(* IEC 61131-3 sources: plcassist-cli/packages/volt-lsp-iec/test-corpus/lenze-mid/Device/Plc Logic/Application/A70_MachineModuleSources/MM_MachineControl/01_Main, 9 files *)

(* ---- Mach1_Drives.fb ---- *)
FUNCTION_BLOCK Mach1_Drives
VAR_INPUT
END_VAR
VAR_OUTPUT
END_VAR
VAR
	testbyte: BYTE;
	testdint: DWORD;
	testword: WORD;
	OspRotationFlag: R_TRIG;
	OffDelayEnableDrivePower: TOF;
	EnableDrivePower: BOOL;
	bServoDrivesInSync: BOOL;
	TimeOutInSync: TON;
	bInSyncTimeOut: BOOL;
	TimeOutInLock: TON;
	tSetDrivesInLock: BOOL;
	bInLockTimeOut: BOOL;
	SideCorrection_CW: sUDT_ServoComm_Drive_Control;
	Servo_LimitJog_Instance: Servo_LimitJog;
	FBFeedforwardADS: FB_Lenze_i550;
	FBFeedforwardATF: FB_Lenze_i550;
	FBElevatorATF: FB_Lenze_i550;
	FBFan: FB_Lenze_i550;
	FBBobbin: FB_Lenze_i550;
	tReal: REAL;
	tWrapperStopPosition: DINT;

	sadad: FB_Lenze_i550;
	FB_Lenze_i550_0: FB_Lenze_i550;

mydword:DWORD;

	tbool: BOOL;
	OnDelayEnableSync: TON;
	ScaleBobbinTorque: LIN_TRAFO;
	tBobbinTorque: REAL;
	OffDelaySync: TOF;
	TON_0: TON;

	MainDrive_VirtualMasterControl: VirtualMasterControl;
END_VAR

VAR CONSTANT
	ctCurveIsSpeed: INT := 2;
	ctCurveIs0ToMax: INT := 0;
END_VAR
VAR
	ServoMainDrive: ServoControl;
	ServoWrappingDevice: ServoControl;
	ServoSideCorrection: ServoControl;
END_VAR

NETWORK 0 LD TITLE: "DONE network 3 : All drives ready"
  Mach1.GenFlags.ConditionsReadyForOperation := ((Mach1_Data.Drives.MainDrive.Status.DriveIsReady OR NOT Mach1_Data.Drives.MainDrive.Control.SetDriveEnable) AND (Mach1_Data.Drives.WrappingDevice.Status.DriveIsReady OR NOT Mach1_Data.Drives.WrappingDevice.Control.SetDriveEnable) AND (Mach1_Data.Drives.SideCorrection.Status.DriveIsReady OR NOT Mach1_Data.Drives.SideCorrection.Control.SetDriveEnable));
END_NETWORK
NETWORK 1 LD
  LET g24 := EnableDrivePower;
  Mach1_Data.Drives.WrappingDevice.Control.StartSetHomePos R= (g24 AND Mach1_Data.Drives.WrappingDevice.Status.DriveIsHomed);
  Mach1_Data.Drives.WrappingDevice.Control.StartSetHomePos S= ((g24 AND NOT Mach1_Data.Drives.WrappingDevice.Status.DriveIsHomed) AND FF500ms);
END_NETWORK
NETWORK 2 LD TITLE: "DONE Network 4: Enable drive power"
  // The off delay ensures that the drive can stop before the power is removed from the drive. The power must be removed from the drive before it goes to STO. If the power remains on during STO, the drive will generate an error.
  EnableDrivePower := (TRUE AND Mach1_Safety.Status.STO_OK);
END_NETWORK
NETWORK 3 LD
  Mach1_AuxData.AllDrivesHomed := Mach1_Data.Drives.MainDrive.Status.DriveIsHomed;
END_NETWORK
NETWORK 4 LD
  LET g0 := TRUE;
  Mach1_Data.Drives.MainDrive_VM.Control.SetDriveEnable := (g0 AND mach1.Genflags.DelayAfterSTO);
  Mach1_Data.Drives.MainDrive_VM.Control.ResetError := ((g0 AND NOT Mach1_Data.Drives.MainDrive_VM.Status.DriveIsReady) AND FF100ms);
  LET en1 := g0;
  IF en1 THEN MainDrive_VirtualMasterControl(iAcc := 600, iDec := 1800, ioVirtualMaster := Mach1_Data.Drives.MainDrive_VM, ioVirtualMasterCom := Data_Exchange_Motion.Servo_VirtualMaster); END_IF
  LET en2 := g0;
  IF en2 THEN HMI_Var.Mach1.ActualSpeed := MOVE(Mach1_Data.Drives.MainDrive_VM.Status.ActSpeed); END_IF
  LET en3 := en2;
  IF en3 THEN HMI_Var.Mach1.Position := MOVE(Mach1_Data.Drives.MainDrive_VM.Status.ActXPos); END_IF
END_NETWORK
NETWORK 5 LD TITLE: "Warning: machine in manual homing mode"
  Alarms_V5_1_100(Mach1_Alarms, (Mach1.GenFlags.DelayAfterSTO AND Mach1_AuxData.EnableManualHomeSetting), Mach1.GenFlags.ResetFlag, Mach1_Alarms.Alm033, Mach1.GenFlags.Warning);
END_NETWORK
NETWORK 6 LD TITLE: "DONE Network 5 : Conditions for sync/lock"
  LET g1 := Mach1.GenFlags.DelayAfterEmergStop;
  Mach1_AuxData.SetDrivesInSync := (TON_0(IN := (OffDelaySync(IN := (g1 AND Mach1_Safety.Status.DoorsOK), PT := T#500MS) AND Mach1_Safety.Status.STO_OK), PT := T#500MS) AND Mach1.GenFlags.ConditionsReadyForOperation AND Mach1_AuxData.AllDrivesHomed AND NOT Mach1_AuxData.EnableManualHomeSetting);
  LET g2 := (g1 AND Mach1_AuxData.SetDrivesInSync);
  bServoDrivesInSync := (g2 AND Mach1_Data.Drives.MainDrive.Status.InSync AND (Mach1_Data.Drives.WrappingDevice.Status.InSync OR NOT Mach1_Data.Drives.WrappingDevice.Control.SetDriveEnable) AND (Mach1_Data.Drives.SideCorrection.Status.InSync OR NOT Mach1_Data.Drives.SideCorrection.Control.SetDriveEnable));
  bInSyncTimeOut := TimeOutInSync(IN := (g2 AND NOT bServoDrivesInSync), PT := T#10S);
  Mach1_AuxData.SetDrivesInLock := ((g1 AND bServoDrivesInSync) AND (Mach1_AuxData.IEC_TIMERS.OffDelayLockDrives(IN := , PT := T#2s) OR TRUE));
  LET g3 := (g1 AND (Mach1_AuxData.SetDrivesInLock OR Mach1_AuxData.SetDrivesInSync));
  Mach1_AuxData.AllDrivesInLock := (g3 AND Mach1_Data.Drives.MainDrive.Status.InSync AND (Mach1_Data.Drives.WrappingDevice.Status.InSync OR NOT Mach1_Data.Drives.WrappingDevice.Control.SetDriveEnable) AND (Mach1_Data.Drives.SideCorrection.Status.InSync OR NOT Mach1_Data.Drives.SideCorrection.Control.SetDriveEnable));
  bInLockTimeOut := TimeOutInLock(IN := (g3 AND NOT Mach1_AuxData.AllDrivesInLock), PT := T#5S);
  tSetDrivesInLock := g3;
END_NETWORK
NETWORK 7 LD TITLE: "DONE Network 6: Servo Main drive: Control"
  LET g4 := TRUE;
  Mach1_Data.Drives.MainDrive_VM.Control.StartMovement := (g4 AND ((Mach1_Safety.Control.RequestManSpeed AND Mach1_Safety.Status.SafetyManSpeed) OR (Mach1_Safety.Control.RequestAutoSpeed AND Mach1_Safety.Status.SafetyAutoSpeed)));
  LET en1 := (g4 AND TRUE);
  IF en1 THEN Mach1_Data.Drives.MainDrive.CAM.CamType := MOVE(ctCurveIs0ToMax); END_IF
  Mach1_Data.Drives.MainDrive.Control.SetInSync := (en1 AND tSetDrivesInLock);
  LET g5 := (g4 AND TRUE);
  Mach1_Data.Drives.MainDrive.Control.SetBrakeRelease := (g5 AND Mach1_Alarms.Alm001 AND HMI_Var.ReleaseBrake);
  HMI_Var.ReleaseBrake R= (g5 AND (NOT Mach1_Alarms.Alm001 OR (mach1.Genflags.StartFlag AND Mach1_Alarms.Alm001)));
  LET en2 := (g4 AND TRUE);
  IF en2 THEN ServoMainDrive(iServoStatus := Data_Exchange_Motion.Servo_MainDrive.Status, iEnableHomeMovement := TRUE, iEnablePower := EnableDrivePower, iFF100ms := LST_General.FF100ms, ioUDT_ServoDrive := Mach1_Data.Drives.MainDrive, oServoControl => Data_Exchange_Motion.Servo_MainDrive.Control); END_IF
  Mach1.GenFlags.Rotflag := OspRotationFlag(CLK := (en2 AND Mach1_Data.Drives.MainDrive.Status.RotationPulse));
END_NETWORK
NETWORK 8 LD TITLE: "DONE Network 7 : Servo Main drive: Alarms"
  Mach1.GenFlags.StopDriveDirect S= (Alarms_V5_1_100(Mach1_Alarms, (Mach1.GenFlags.DelayAfterSTO AND NOT Mach1_Data.Drives.MainDrive.Status.DriveIsReady), Mach1.GenFlags.ResetFlag, Mach1_Alarms.Alm020, Mach1.GenFlags.MinorAlarm) OR Alarms_V5_1_100(Mach1_Alarms, (Mach1.GenFlags.DelayAfterSTO AND Mach1_Data.Drives.MainDrive.Status.DriveTorqueError), Mach1.GenFlags.ResetFlag, Mach1_Alarms.Alm021, Mach1.GenFlags.MinorAlarm) OR Alarms_V5_1_100(Mach1_Alarms, (Mach1.GenFlags.DelayAfterSTO AND NOT Mach1_Data.Drives.MainDrive.Status.DriveIsHomed), Mach1.GenFlags.ResetFlag, Mach1_Alarms.Alm022, Mach1.GenFlags.MinorAlarm));
END_NETWORK
NETWORK 9 LD
  Mach1_Data.Drives.MainDrive.Control.ResetError S= (((Mach1_Alarms.Alm020 OR Mach1_Alarms.Alm021 OR Mach1_Alarms.Alm022) AND Mach1.GenFlags.ResetFlag) OR (TON_0.Q AND Imp100ms AND Mach1_Safety.Status.ServiceMode AND Mach1_Safety.Status.Service_ButtonAB));
END_NETWORK
NETWORK 10 LD TITLE: "DONE Network 8: Servo Wrapping device: Control"
  LET g6 := TRUE;
  LET en1 := (g6 AND TRUE);
  IF en1 THEN Mach1_Data.Drives.WrappingDevice.CAM.CamType := MOVE(ctCurveIsSpeed); END_IF
  Mach1_Data.Drives.WrappingDevice.Control.SetInSync := (en1 AND tSetDrivesInLock);
  LET en2 := g6;
  IF en2 THEN Mach1_Data.Drives.WrappingDevice.CAM.Y_Scale_Recipe := MOVE(Mach1_Data.Settings.Ints.RollingDeviceSpeedFactor); END_IF
  LET en3 := (g6 AND TRUE);
  IF en3 THEN ServoWrappingDevice(iServoStatus := Data_Exchange_Motion.Servo_WrappingDevice.Status, iEnableHomeMovement := TRUE, iEnablePower := EnableDrivePower, iFF100ms := LST_General.FF100ms, ioUDT_ServoDrive := Mach1_Data.Drives.WrappingDevice, oServoControl => Data_Exchange_Motion.Servo_WrappingDevice.Control); END_IF
END_NETWORK
NETWORK 11 LD TITLE: "DONE Network 9 : Servo Wrapping Device: Alarms"
  LET g7 := (Alarms_V5_1_100(Mach1_Alarms, (Mach1.GenFlags.DelayAfterSTO AND NOT Mach1_Data.Drives.WrappingDevice.Status.DriveIsReady AND Mach1_Data.Drives.WrappingDevice.Control.SetDriveEnable), Mach1.GenFlags.ResetFlag, Mach1_Alarms.Alm023, Mach1.GenFlags.MinorAlarm) OR Alarms_V5_1_100(Mach1_Alarms, (Mach1.GenFlags.DelayAfterSTO AND Mach1_Data.Drives.WrappingDevice.Status.DriveTorqueError), Mach1.GenFlags.ResetFlag, Mach1_Alarms.Alm024, Mach1.GenFlags.MinorAlarm) OR Alarms_V5_1_100(Mach1_Alarms, (Mach1.GenFlags.DelayAfterSTO AND NOT Mach1_Data.Drives.WrappingDevice.Status.DriveIsHomed), Mach1.GenFlags.ResetFlag, Mach1_Alarms.Alm025, Mach1.GenFlags.MinorAlarm));
  Mach1.GenFlags.StopDriveDirect S= g7;
  Mach1_Data.Drives.WrappingDevice.Control.ResetError S= (g7 AND Mach1.GenFlags.ResetFlag);
END_NETWORK
NETWORK 12 LD
  Mach1_Data.Drives.WrappingDevice.Control.ResetError S= (((Mach1_Alarms.Alm023 OR Mach1_Alarms.Alm024 OR Mach1_Alarms.Alm025) AND Mach1.GenFlags.ResetFlag) OR (TON_0.Q AND Imp100ms AND Mach1_Safety.Status.ServiceMode AND Mach1_Safety.Status.Service_ButtonAB));
END_NETWORK
NETWORK 13 LD
END_NETWORK
NETWORK 14 LD TITLE: "Digital inputs"
  // 16: non-motor side
  // 17: motor side
  LET en1 := TRUE;
  IF en1 THEN mydword := MOVE(%ID79); END_IF
  LET g8 := en1;
  Data_Exchange_Motion.Servo_SideCorrection.Status.Spare1 := (g8 AND mydword.16);
  Data_Exchange_Motion.Servo_SideCorrection.Status.Spare2 := (g8 AND mydword.17);
END_NETWORK
NETWORK 15 LD TITLE: "DONE Network 10: Servo Side correction: Control"
  LET g9 := TRUE;
  LET en1 := (g9 AND TRUE);
  IF en1 THEN Mach1_Data.Drives.SideCorrection.CAM.CamType := MOVE(ctCurveIsSpeed); END_IF
  Mach1_Data.Drives.SideCorrection.Control.SetInSync := (en1 AND tSetDrivesInLock);
  LET en2 := (g9 AND TRUE);
  IF en2 THEN ServoSideCorrection(iServoStatus := Data_Exchange_Motion.Servo_SideCorrection.Status, iEnableHomeMovement := TRUE, iEnablePower := EnableDrivePower, iFF100ms := LST_General.FF100ms, ioUDT_ServoDrive := Mach1_Data.Drives.SideCorrection, oServoControl => SideCorrection_CW); END_IF
  LET en3 := (g9 AND TRUE);
  IF en3 THEN Servo_LimitJog_Instance(iServoStatus := Data_Exchange_Motion.Servo_SideCorrection.Status, iServoControl := SideCorrection_CW, ioUDT_ServoDrive := Mach1_Data.Drives.SideCorrection, ioUDT_JogLimitFree := Mach1_Data.Drives.SideCorrection_FreeLimit, oServoControl => Data_Exchange_Motion.Servo_SideCorrection.Control); END_IF
END_NETWORK
NETWORK 16 LD TITLE: "DONE Network 11 : Servo Side correction: Alarms"
  LET g10 := (Alarms_V5_1_100(Mach1_Alarms, (Mach1.GenFlags.DelayAfterSTO AND NOT Mach1_Data.Drives.SideCorrection.Status.DriveIsReady AND Mach1_Data.Drives.SideCorrection.Control.SetDriveEnable), Mach1.GenFlags.ResetFlag, Mach1_Alarms.Alm026, Mach1.GenFlags.MinorAlarm) OR Alarms_V5_1_100(Mach1_Alarms, (Mach1.GenFlags.DelayAfterSTO AND Mach1_Data.Drives.SideCorrection.Status.DriveTorqueError), Mach1.GenFlags.ResetFlag, Mach1_Alarms.Alm027, Mach1.GenFlags.MinorAlarm) OR Alarms_V5_1_100(Mach1_Alarms, (Mach1.GenFlags.DelayAfterSTO AND NOT Mach1_Data.Drives.SideCorrection.Status.DriveIsHomed), Mach1.GenFlags.ResetFlag, Mach1_Alarms.Alm028, Mach1.GenFlags.MinorAlarm));
  Mach1.GenFlags.StopDriveDirect S= g10;
  Mach1_Data.Drives.SideCorrection.Control.ResetError S= (g10 AND Mach1.GenFlags.ResetFlag);
END_NETWORK
NETWORK 17 LD
  Mach1_Data.Drives.SideCorrection.Control.ResetError S= (((Mach1_Alarms.Alm026 OR Mach1_Alarms.Alm027 OR Mach1_Alarms.Alm028) AND Mach1.GenFlags.ResetFlag) OR (TON_0.Q AND Imp100ms AND Mach1_Safety.Status.ServiceMode AND Mach1_Safety.Status.Service_ButtonAB));
END_NETWORK
NETWORK 18 LD
END_NETWORK
NETWORK 19 LD TITLE: "DONE Network 12: Feedforward ADS"
  LET g11 := TRUE;
  Mach1_Data.Drives.FeedForwardADS.Control.Enable := (g11 AND Mach1.GenFlags.DelayAfterEmergStop AND NOT Mach1_Alarms.Alm015);
  Mach1_Data.Drives.FeedForwardADS.Control.Reverse := g11;
  LET en1 := g11;
  IF en1 THEN FBFeedforwardADS(iStatusWord := Data_Exchange_Motion.FQI_FeedforwardADS.Status, iGearRatioNumerator := 2790.0, iGearRatioDenominator := 111.0, iNominalMotorSpeedwoSlipComp_RPM := 3000.0, iNominalMotorFrequency_Hz := 100.0, iAxisJogSpeed_RPM := 10.0, ioUDT := Mach1_Data.Drives.FeedForwardADS, oControlWord => Data_Exchange_Motion.FQI_FeedforwardADS.Controlword, oRefSpeed => Data_Exchange_Motion.FQI_FeedforwardADS.RefSpeed); END_IF
END_NETWORK
NETWORK 20 LD TITLE: "DONE Network 13: Alarms feed forward dryer"
  LET g12 := Alarms_V5_1_100(Mach1_Alarms, (Mach1.GenFlags.DelayAfterEmergStop AND Mach1_Data.Drives.FeedForwardADS.Status.Error), True, Mach1_Alarms.Alm015, Mach1.GenFlags.MinorAlarm);
  Mach1.GenFlags.StopDriveDirect S= g12;
  Mach1_Data.Drives.FeedForwardADS.Control.ResetError S= (g12 AND Mach1.GenFlags.ResetFlag);
END_NETWORK
NETWORK 21 LD TITLE: "DONE Network 14: Feedforward ATF"
  LET g13 := TRUE;
  Mach1_Data.Drives.FeedForwardATF.Control.Enable := (g13 AND Mach1.GenFlags.DelayAfterEmergStop AND NOT Mach1_Alarms.Alm016);
  LET en1 := g13;
  IF en1 THEN FBFeedforwardATF(iStatusWord := Data_Exchange_Motion.FQI_FeedforwardATF.Status, iGearRatioNumerator := 2790.0, iGearRatioDenominator := 111.0, iNominalMotorSpeedwoSlipComp_RPM := 3000.0, iNominalMotorFrequency_Hz := 100.0, iAxisJogSpeed_RPM := 10.0, ioUDT := Mach1_Data.Drives.FeedForwardATF, oControlWord => Data_Exchange_Motion.FQI_FeedforwardATF.Controlword, oRefSpeed => Data_Exchange_Motion.FQI_FeedforwardATF.RefSpeed); END_IF
END_NETWORK
NETWORK 22 LD TITLE: "DONE Network 15: Alarms feed forward trayfiller"
  LET g14 := Alarms_V5_1_100(Mach1_Alarms, (Mach1.GenFlags.DelayAfterEmergStop AND Mach1_Data.Drives.FeedForwardATF.Status.Error), True, Mach1_Alarms.Alm016, Mach1.GenFlags.MinorAlarm);
  Mach1.GenFlags.StopDriveDirect S= g14;
  Mach1_Data.Drives.FeedForwardATF.Control.ResetError S= (g14 AND Mach1.GenFlags.ResetFlag);
END_NETWORK
NETWORK 23 LD TITLE: "DONE Network 16: Elevator ATF"
  LET g15 := TRUE;
  Mach1_Data.Drives.ElevatorATF.Control.Enable := (g15 AND Mach1.GenFlags.DelayAfterEmergStop AND NOT Mach1_Alarms.Alm014);
  LET en1 := g15;
  IF en1 THEN FBElevatorATF(iStatusWord := Data_Exchange_Motion.FQI_ElevatorATF.Status, iGearRatioNumerator := 100.0, iGearRatioDenominator := 111.0, iNominalMotorSpeedwoSlipComp_RPM := 3000.0, iNominalMotorFrequency_Hz := 100.0, iAxisJogSpeed_RPM := 10.0, ioUDT := Mach1_Data.Drives.ElevatorATF, oControlWord => Data_Exchange_Motion.FQI_ElevatorATF.Controlword, oRefSpeed => Data_Exchange_Motion.FQI_ElevatorATF.RefSpeed); END_IF
END_NETWORK
NETWORK 24 LD TITLE: "DONE Network 17: Alarms Elevator trayfiller"
  LET g16 := Alarms_V5_1_100(Mach1_Alarms, (Mach1.GenFlags.DelayAfterEmergStop AND Mach1_Data.Drives.ElevatorATF.Status.Error), True, Mach1_Alarms.Alm014, Mach1.GenFlags.MinorAlarm);
  Mach1.GenFlags.StopDriveDirect S= g16;
  Mach1_Data.Drives.ElevatorATF.Control.ResetError S= (g16 AND Mach1.GenFlags.ResetFlag);
END_NETWORK
NETWORK 25 LD TITLE: "DONE Network 18: Fan"
  LET g26 := TRUE;
  Mach1_Data.Drives.Fan.Control.Enable := (g26 AND Mach1.GenFlags.EnableAuxDrive AND NOT Mach1_Alarms.Alm017);
  LET en1 := g26;
  IF en1 THEN FBFan(iStatusWord := Data_Exchange_Motion.FQI_Fan.Status, iGearRatioNumerator := 1.0, iGearRatioDenominator := 1.0, iNominalMotorSpeedwoSlipComp_RPM := 3000.0, iNominalMotorFrequency_Hz := 50.0, iAxisJogSpeed_RPM := 10.0, ioUDT := Mach1_Data.Drives.Fan, oControlWord => Data_Exchange_Motion.FQI_Fan.Controlword, oRefSpeed => Data_Exchange_Motion.FQI_Fan.RefSpeed); END_IF
END_NETWORK
NETWORK 26 LD TITLE: "DONE Network 19: Alarms Fan"
  LET g18 := Alarms_V5_1_100(Mach1_Alarms, (Mach1.GenFlags.DelayAfterEmergStop AND Mach1_Data.Drives.Fan.Status.Error), True, Mach1_Alarms.Alm017, Mach1.GenFlags.MinorAlarm);
  Mach1.GenFlags.StopDriveDirect S= g18;
  Mach1_Data.Drives.Fan.Control.ResetError S= (g18 AND Mach1.GenFlags.ResetFlag);
END_NETWORK
NETWORK 27 LD TITLE: "DONE Network 20: Bobbin"
  LET g19 := TRUE;
  LET en1 := (g19 AND Mach1.GenFlags.EnableAuxDrive AND NOT HMI_Var.Btn_Cleaning);
  IF en1 THEN (Mach1_Data.Settings.Ints.TorqueControlBobbin > 0); END_IF
  LET g20 := (en1 AND Mach1_Safety.Status.AllDoorsActuallyClosed);
  Mach1_Data.Drives.Bobbine.Control.Enable := g20;
  LET en2 := g20;
  IF en2 THEN Mach1_Data.Drives.Bobbine.Control.AutoSpeed := MOVE(860); END_IF
  Mach1_Data.Drives.Bobbine.Control.StartAuto := en2;
  LET en3 := g19;
  IF en3 THEN FBBobbin(iStatusWord := Data_Exchange_Motion.FQI_Bobbin.Status, iGearRatioNumerator := 2790.0, iGearRatioDenominator := 111.0, iNominalMotorSpeedwoSlipComp_RPM := 3000.0, iNominalMotorFrequency_Hz := 50.0, iAxisJogSpeed_RPM := 10.0, ioUDT := Mach1_Data.Drives.Bobbine, oControlWord => Data_Exchange_Motion.FQI_Bobbin.Controlword, oRefSpeed => Data_Exchange_Motion.FQI_Bobbin.RefSpeed); END_IF
  LET g21 := (g19 AND HMI_Var.Mach1.CalibrateTorqueValues);
  LET en4 := g21;
  IF en4 THEN Data_Exchange_Motion.BobbinTorque := MOVE(Mach1_AuxData.TorqueCalibrationValue); END_IF
  LET en5 := (g21 AND HMI_Var.Mach1.setMinTorqueValue);
  IF en5 THEN Mach1_Data.Settings.Dints.minTorqueValue := MOVE(Mach1_AuxData.TorqueCalibrationValue); END_IF
  HMI_Var.Mach1.setMinTorqueValue R= en5;
  LET en6 := (g21 AND HMI_Var.Mach1.setMaxTorqueValue);
  IF en6 THEN Mach1_Data.Settings.Dints.maxTorqueValue := MOVE(Mach1_AuxData.TorqueCalibrationValue); END_IF
  HMI_Var.Mach1.setMaxTorqueValue R= en6;
  LET i1 := DINT_TO_REAL(Mach1_Data.Settings.Dints.minTorqueValue);
  LET i2 := DINT_TO_REAL(Mach1_Data.Settings.Dints.maxTorqueValue);
  LET en7 := (g19 AND NOT HMI_Var.Mach1.CalibrateTorqueValues);
  IF en7 THEN ScaleBobbinTorque(IN := Mach1_Data.Settings.Ints.TorqueControlBobbin, IN_MIN := 0, IN_MAX := 1000, OUT_MIN := i1, OUT_MAX := i2, OUT => tBobbinTorque); END_IF
  LET i3 := REAL_TO_DINT(tBobbinTorque);
  LET en8 := en7;
  IF en8 THEN Data_Exchange_Motion.BobbinTorque := MOVE(i3); END_IF
END_NETWORK
NETWORK 28 LD TITLE: "DONE Network 21: Alarms Bobbine"
  LET g22 := Alarms_V5_1_100(Mach1_Alarms, (Mach1_AuxData.MIDS_Active AND Mach1.GenFlags.DelayAfterEmergStop AND NOT Mach1_Data.Drives.Bobbine.Status.DriveReady AND Mach1_AuxData.AllDrivesHomed), True, Mach1_Alarms.Alm010, Mach1.GenFlags.MinorAlarm);
  Mach1.GenFlags.StopDriveDirect S= g22;
  Mach1_Data.Drives.Bobbine.Control.ResetError S= (g22 AND Mach1.GenFlags.ResetFlag);
END_NETWORK
NETWORK 29 LD TITLE: "TODO Network 22:"
  // WRAPPER
END_NETWORK
NETWORK 30 LD TITLE: "TODO Network 23: Limit Wrapper stop position"
  LET g23 := TRUE;
  LET en1 := g23;
  IF en1 THEN (Mach1_Data.Settings.Dints.WrapperStopPosition > 400); END_IF
  LET en2 := en1;
  IF en2 THEN Mach1_Data.Settings.Dints.WrapperStopPosition := MOVE(400); END_IF
  LET en3 := g23;
  IF en3 THEN (Mach1_Data.Settings.Dints.WrapperStopPosition < 5); END_IF
  LET en4 := en3;
  IF en4 THEN Mach1_Data.Settings.Dints.WrapperStopPosition := MOVE(5); END_IF
  LET en5 := g23;
  IF en5 THEN tWrapperStopPosition := (Mach1_Data.Settings.Dints.WrapperStopPosition * 100); END_IF
END_NETWORK
NETWORK 31 LD TITLE: "TODO Network 25:"
  Data_Exchange_Motion.FeedForwardWrapper.Control.Enable := (TRUE AND Mach1.GenFlags.DelayAfterEmergStop AND NOT Mach1_Alarms.Alm066);
END_NETWORK
NETWORK 32 LD TITLE: "TODO Network 26:"
  LET g1 := (Alarms_V5_1_100(Mach1_Alarms, (Mach1_AuxData.MIDS_Active AND Mach1.GenFlags.EnableMainDrive AND HMI_Var.Test_Prod AND NOT HMI_Var.Btn_Cleaning AND Mach1_AuxData.AllDrivesHomed AND NOT Data_Exchange_Motion.FeedForwardWrapper.Status.ReadyForMotion), Mach1.Genflags.StartFlag, Mach1_Alarms.Alm056, Mach1.GenFlags.MinorAlarm) AND mach1.Genflags.ResetFlag);
  Mach1_Data.Drives.WrappingDevice.Control.ResetError S= g1;
  Data_Exchange_Motion.FeedForwardWrapper.Control.ResetError := g1;
END_NETWORK
NETWORK 33 LD TITLE: "TODO Network 27:"
  ;
END_NETWORK

END_FUNCTION_BLOCK

(* ---- fc_Information.prg ---- *)
PROGRAM fc_Information
VAR
END_VAR

VersionInfo_DB.PLC_version:='MID-S100-L-V00_00';
VersionInfo_DB.PLC_Version_Date:='08-06-2023';

END_PROGRAM

(* ---- ForceOutput.prg ---- *)
PROGRAM ForceOutput
VAR
END_VAR

NETWORK 0 LD
  LET g2 := HMI_Var.ForceOutputs;
  LST_InputsOutputs.Q100_0_Pilot_light_Alarm_green_ := (g2 AND LST_InputsOutputs.Serv_QB100.0);
  LST_InputsOutputs.Q100_1_Pilot_light_Alarm_orange_ := (g2 AND LST_InputsOutputs.Serv_QB100.1);
  LST_InputsOutputs.Q100_2_Pilot_light_Alarm_red_ := (g2 AND LST_InputsOutputs.Serv_QB100.2);
  LST_InputsOutputs.Q100_3_Pilot_light_Alarm_buzzer_ := (g2 AND LST_InputsOutputs.Serv_QB100.3);
  LST_InputsOutputs.Q100_4_Spare := (g2 AND LST_InputsOutputs.Serv_QB100.4);
  LST_InputsOutputs.Q100_5_Signal_lamp_Start := (g2 AND LST_InputsOutputs.Serv_QB100.5);
  LST_InputsOutputs.Q100_6_Signal_lamp_Stop := (g2 AND LST_InputsOutputs.Serv_QB100.6);
  LST_InputsOutputs.Q100_7_Activate_greasing_system := (g2 AND LST_InputsOutputs.Serv_QB100.7);
  LST_InputsOutputs.Q101_0_REL_release_brake := (g2 AND LST_InputsOutputs.Serv_QB101.0);
  LST_InputsOutputs.Q101_1_PNV_Waterlevel_control := (g2 AND LST_InputsOutputs.Serv_QB101.1);
  LST_InputsOutputs.Q101_2_Enable_GluePump := (g2 AND LST_InputsOutputs.Serv_QB101.2);
  LST_InputsOutputs.Q101_3_Spare := (g2 AND LST_InputsOutputs.Serv_QB101.3);
  LST_InputsOutputs.Q101_4_Spare := (g2 AND LST_InputsOutputs.Serv_QB101.4);
  LST_InputsOutputs.Q101_5_Spare := (g2 AND LST_InputsOutputs.Serv_QB101.5);
  LST_InputsOutputs.Q101_6_Spare := (g2 AND LST_InputsOutputs.Serv_QB101.6);
  LST_InputsOutputs.Q101_7_Spare := (g2 AND LST_InputsOutputs.Serv_QB101.7);
END_NETWORK
NETWORK 1 LD
  LET g1 := HMI_Var.ForceOutputs;
  LST_InputsOutputs.Q132_0_SL_Start_OP2a := (g1 AND LST_InputsOutputs.Serv_QB132.0);
  LST_InputsOutputs.Q132_1_SL_Stop_OP2a := (g1 AND LST_InputsOutputs.Serv_QB132.1);
  LST_InputsOutputs.Q132_2_Enable_power_controllers := (g1 AND LST_InputsOutputs.Serv_QB132.2);
  LST_InputsOutputs.Q132_3_Spare := (g1 AND LST_InputsOutputs.Serv_QB132.3);
  LST_InputsOutputs.Q132_4_CT_Fan_dryer := (g1 AND LST_InputsOutputs.Serv_QB132.4);
  LST_InputsOutputs.Q132_5_Spare := (g1 AND LST_InputsOutputs.Serv_QB132.5);
  LST_InputsOutputs.Q132_6_PNV_Inpusher := (g1 AND LST_InputsOutputs.Serv_QB132.6);
  LST_InputsOutputs.Q132_7_PNV_tilting_inpusher := (g1 AND LST_InputsOutputs.Serv_QB132.7);
  LST_InputsOutputs.Q133_0_Spare := (g1 AND LST_InputsOutputs.Serv_QB133.0);
  LST_InputsOutputs.Q133_1_Spare := (g1 AND LST_InputsOutputs.Serv_QB133.1);
  LST_InputsOutputs.Q133_2_Spare := (g1 AND LST_InputsOutputs.Serv_QB133.2);
  LST_InputsOutputs.Q133_3_Spare := (g1 AND LST_InputsOutputs.Serv_QB133.3);
  LST_InputsOutputs.Q133_4_Spare := (g1 AND LST_InputsOutputs.Serv_QB133.4);
  LST_InputsOutputs.Q133_5_InfeedConv_Fwd := (g1 AND LST_InputsOutputs.Serv_QB133.5);
  LST_InputsOutputs.Q133_6_InfeedConv_Rev := (g1 AND LST_InputsOutputs.Serv_QB133.6);
  LST_InputsOutputs.Q133_7_OutfeedConv_Fwd := (g1 AND LST_InputsOutputs.Serv_QB133.7);
END_NETWORK
NETWORK 2 LD
  LET g0 := HMI_Var.ForceOutputs;
  LST_InputsOutputs.Q136_0_Spare := (g0 AND LST_InputsOutputs.Serv_QB136.0);
  LST_InputsOutputs.Q136_1_Spare := (g0 AND LST_InputsOutputs.Serv_QB136.1);
  LST_InputsOutputs.Q136_2_Spare := (g0 AND LST_InputsOutputs.Serv_QB136.2);
  LST_InputsOutputs.Q136_3_Spare := (g0 AND LST_InputsOutputs.Serv_QB136.3);
  LST_InputsOutputs.Q136_4_Spare := (g0 AND LST_InputsOutputs.Serv_QB136.4);
  LST_InputsOutputs.Q136_5_Spare := (g0 AND LST_InputsOutputs.Serv_QB136.5);
  LST_InputsOutputs.Q136_6_Spare := (g0 AND LST_InputsOutputs.Serv_QB136.6);
  LST_InputsOutputs.Q136_7_Spare := (g0 AND LST_InputsOutputs.Serv_QB132.7);
  LST_InputsOutputs.Q137_0_Spare := (g0 AND LST_InputsOutputs.Serv_QB137.0);
  LST_InputsOutputs.Q137_1_Spare := (g0 AND LST_InputsOutputs.Serv_QB137.1);
  LST_InputsOutputs.Q137_2_Spare := (g0 AND LST_InputsOutputs.Serv_QB137.2);
  LST_InputsOutputs.Q137_3_Spare := (g0 AND LST_InputsOutputs.Serv_QB137.3);
  LST_InputsOutputs.Q137_4_Spare := (g0 AND LST_InputsOutputs.Serv_QB137.4);
  LST_InputsOutputs.Q137_5_Spare := (g0 AND LST_InputsOutputs.Serv_QB137.5);
  LST_InputsOutputs.Q137_6_Spare := (g0 AND LST_InputsOutputs.Serv_QB137.6);
  LST_InputsOutputs.Q137_7_Spare := (g0 AND LST_InputsOutputs.Serv_QB137.7);
END_NETWORK
NETWORK 3 LD
END_NETWORK

END_PROGRAM

(* ---- ForceOutput_1.prg ---- *)
PROGRAM ForceOutput_1
VAR
END_VAR

NETWORK 0 LD
  LET g2 := NOT HMI_Var.ForceOutputs;
  LST_InputsOutputs.Serv_QB100.0 := (g2 AND LST_InputsOutputs.Q100_0_Pilot_light_Alarm_green_);
  LST_InputsOutputs.Serv_QB100.1 := (g2 AND LST_InputsOutputs.Q100_1_Pilot_light_Alarm_orange_);
  LST_InputsOutputs.Serv_QB100.2 := (g2 AND LST_InputsOutputs.Q100_2_Pilot_light_Alarm_red_);
  LST_InputsOutputs.Serv_QB100.3 := (g2 AND LST_InputsOutputs.Q100_3_Pilot_light_Alarm_buzzer_);
  LST_InputsOutputs.Serv_QB100.4 := (g2 AND LST_InputsOutputs.Q100_4_Spare);
  LST_InputsOutputs.Serv_QB100.5 := (g2 AND LST_InputsOutputs.Q100_5_Signal_lamp_Start);
  LST_InputsOutputs.Serv_QB100.6 := (g2 AND LST_InputsOutputs.Q100_6_Signal_lamp_Stop);
  LST_InputsOutputs.Serv_QB100.7 := (g2 AND LST_InputsOutputs.Q100_7_Activate_greasing_system);
  LST_InputsOutputs.Serv_QB101.0 := (g2 AND LST_InputsOutputs.Q101_0_REL_release_brake);
  LST_InputsOutputs.Serv_QB101.1 := (g2 AND LST_InputsOutputs.Q101_1_PNV_Waterlevel_control);
  LST_InputsOutputs.Serv_QB101.2 := (g2 AND LST_InputsOutputs.Q101_2_Enable_GluePump);
  LST_InputsOutputs.Serv_QB101.3 := (g2 AND LST_InputsOutputs.Q101_3_Spare);
  LST_InputsOutputs.Serv_QB101.4 := (g2 AND LST_InputsOutputs.Q101_4_Spare);
  LST_InputsOutputs.Serv_QB101.5 := (g2 AND LST_InputsOutputs.Q101_5_Spare);
  LST_InputsOutputs.Serv_QB101.6 := (g2 AND LST_InputsOutputs.Q101_6_Spare);
  LST_InputsOutputs.Serv_QB101.7 := (g2 AND LST_InputsOutputs.Q101_7_Spare);
END_NETWORK
NETWORK 1 LD
  LET g1 := NOT HMI_Var.ForceOutputs;
  LST_InputsOutputs.Serv_QB132.0 := (g1 AND LST_InputsOutputs.Q132_0_SL_Start_OP2a);
  LST_InputsOutputs.Serv_QB132.1 := (g1 AND LST_InputsOutputs.Q132_1_SL_Stop_OP2a);
  LST_InputsOutputs.Serv_QB132.2 := (g1 AND LST_InputsOutputs.Q132_2_Enable_power_controllers);
  LST_InputsOutputs.Serv_QB132.3 := (g1 AND LST_InputsOutputs.Q132_3_Spare);
  LST_InputsOutputs.Serv_QB132.4 := (g1 AND LST_InputsOutputs.Q132_4_CT_Fan_dryer);
  LST_InputsOutputs.Serv_QB132.5 := (g1 AND LST_InputsOutputs.Q132_5_Spare);
  LST_InputsOutputs.Serv_QB132.6 := (g1 AND LST_InputsOutputs.Q132_6_PNV_Inpusher);
  LST_InputsOutputs.Serv_QB132.7 := (g1 AND LST_InputsOutputs.Q132_7_PNV_tilting_inpusher);
  LST_InputsOutputs.Serv_QB133.0 := (g1 AND LST_InputsOutputs.Q133_0_Spare);
  LST_InputsOutputs.Serv_QB133.1 := (g1 AND LST_InputsOutputs.Q133_1_Spare);
  LST_InputsOutputs.Serv_QB133.2 := (g1 AND LST_InputsOutputs.Q133_2_Spare);
  LST_InputsOutputs.Serv_QB133.3 := (g1 AND LST_InputsOutputs.Q133_3_Spare);
  LST_InputsOutputs.Serv_QB133.4 := (g1 AND LST_InputsOutputs.Q133_4_Spare);
  LST_InputsOutputs.Serv_QB133.5 := (g1 AND LST_InputsOutputs.Q133_5_InfeedConv_Fwd);
  LST_InputsOutputs.Serv_QB133.6 := (g1 AND LST_InputsOutputs.Q133_6_InfeedConv_Rev);
  LST_InputsOutputs.Serv_QB133.7 := (g1 AND LST_InputsOutputs.Q133_7_OutfeedConv_Fwd);
END_NETWORK
NETWORK 2 LD
  LET g0 := NOT HMI_Var.ForceOutputs;
  LST_InputsOutputs.Serv_QB136.0 := (g0 AND LST_InputsOutputs.Q136_0_Spare);
  LST_InputsOutputs.Serv_QB136.1 := (g0 AND LST_InputsOutputs.Q136_1_Spare);
  LST_InputsOutputs.Serv_QB136.2 := (g0 AND LST_InputsOutputs.Q136_2_Spare);
  LST_InputsOutputs.Serv_QB136.3 := (g0 AND LST_InputsOutputs.Q136_3_Spare);
  LST_InputsOutputs.Serv_QB136.4 := (g0 AND LST_InputsOutputs.Q136_4_Spare);
  LST_InputsOutputs.Serv_QB136.5 := (g0 AND LST_InputsOutputs.Q136_5_Spare);
  LST_InputsOutputs.Serv_QB136.6 := (g0 AND LST_InputsOutputs.Q136_6_Spare);
  LST_InputsOutputs.Serv_QB132.7 := (g0 AND LST_InputsOutputs.Q136_7_Spare);
  LST_InputsOutputs.Serv_QB137.0 := (g0 AND LST_InputsOutputs.Q137_0_Spare);
  LST_InputsOutputs.Serv_QB137.1 := (g0 AND LST_InputsOutputs.Q137_1_Spare);
  LST_InputsOutputs.Serv_QB137.2 := (g0 AND LST_InputsOutputs.Q137_2_Spare);
  LST_InputsOutputs.Serv_QB137.3 := (g0 AND LST_InputsOutputs.Q137_3_Spare);
  LST_InputsOutputs.Serv_QB137.4 := (g0 AND LST_InputsOutputs.Q137_4_Spare);
  LST_InputsOutputs.Serv_QB137.5 := (g0 AND LST_InputsOutputs.Q137_5_Spare);
  LST_InputsOutputs.Serv_QB137.6 := (g0 AND LST_InputsOutputs.Q137_6_Spare);
  LST_InputsOutputs.Serv_QB137.7 := (g0 AND LST_InputsOutputs.Q137_7_Spare);
END_NETWORK
NETWORK 3 LD
END_NETWORK

END_PROGRAM

(* ---- General.prg ---- *)
PROGRAM General
VAR
	WordConvertor: SafetyPLC_WordsToUDT;
	WordConvertor_v2: SafetyPLC_WordsToUDT_v2;
	test_IW132: Bools_To_Byte;
	Qtest: BYTE;
	ib26: INT;
	tbool: BOOL;
	TON_0: TON;
	TON_1: TON;
	BLINK_0: BLINK;
	restart1: BOOL;
END_VAR

NETWORK 0 LD
  LET en1 := TRUE;
  IF en1 THEN GeneralProgramFlags(); END_IF
END_NETWORK
NETWORK 1 LD
  LET en1 := TRUE;
  IF en1 THEN fc_Information(); END_IF
END_NETWORK
NETWORK 2 LD
  WordConvertor_v2(ioSafetyStatusUDT := Mach1_Safety.Status, ioSafetyControlUDT := Mach1_Safety.Control);
END_NETWORK
NETWORK 3 LD
  LET g16 := NOT HMI_Var.ForceOutputs;
  LET en1 := g16;
  IF en1 THEN Mach1_MIDS(); END_IF
  LET en2 := g16;
  IF en2 THEN fc_Visualisation_HMI(); END_IF
  LET en3 := g16;
  IF en3 THEN SMC_BitsToBytes(); END_IF
END_NETWORK
NETWORK 4 LD
  LET en1 := TRUE;
  IF en1 THEN Status_ForceOutputs(); END_IF
END_NETWORK
NETWORK 5 LD
  LST_General.FirstCycle R= ;
END_NETWORK
NETWORK 6 LD
  Bugs.checkconnection := BLINK_0(ENABLE := TRUE, TIMELOW := T#1S, TIMEHIGH := T#1S);
END_NETWORK
NETWORK 7 LD
  TON_0(IN := NOT Bugs.reportConnectionAlive, PT := T#2S);
END_NETWORK
NETWORK 8 LD
  TON_1(IN := Bugs.reportConnectionAlive, PT := T#2S);
END_NETWORK
NETWORK 9 LD
  Bugs.restart := (TON_0.Q OR TON_1.Q);
END_NETWORK

END_PROGRAM

(* ---- Mach1_MIDS.prg ---- *)
PROGRAM Mach1_MIDS
VAR
	FB_Mach1					: GeneralMachineFlags;
	//Mach1.GenFlags				: UDT_GeneralFlags;
	tStopPositionCleaning	: BOOL;

	tDoorUnitOk				: BOOL;
	tCrossDoorcircuit1 		: BOOL;
	tCrossDoorcircuit2 		: BOOL;
	tAlarmlamp				: BOOL;
	tBool					: BOOL;
	tCond					: BOOL;

	tStopPositionLeafCarrier: BOOL;
	tReset: BOOL;
	a:INT;
//TODO
	//test5: CTD;
	//HMI_Var_Mach1_MuteNoBunchAlarm: SR;
	RepetitionNoBunch: CTD;
	tCampulseCigarPresent: BOOL;
	RepetitionNoCigar: CTD;
	PhotocellCigarHasBeenOff: SR;
	tTime1: TIME;
	tLowLevel: BOOL;
	tErrorRuntimeGreasingSystem: BOOL;
	tAlarmSL: BOOL;
	tWarningSL: BOOL;
	tStandbySL: BOOL;
	tRunningSL: BOOL;
	tHeater1Word: WORD;
	tHeater2Word: WORD;
	tHeater3Word: WORD;
	test3: BOOL;
	test4: BOOL;
	qw105: WORD;
	DRYER_SCALING_Heater1: LIN_TRAFO;

	DRYER_Scaling_Speed: LIN_TRAFO;
	lrDryer_ScaledSpeed: REAL;
	lrHeater1_ScaledPower:REAL; //% of max power of 1500

	lrHeater1_Analog: REAL;
	DRYER_SCALING_Heater2: LIN_TRAFO;
	lrHeater2_ScaledPower: REAL;
	DRYER_SCALING_Heater1_Analog: LIN_TRAFO;
	DRYER_SCALING_Heater2_Analog: LIN_TRAFO;
	lrHeater2_Analog: REAL;
	lrHeater3_ScaledPower: REAL;
	DRYER_SCALING_Heater3: LIN_TRAFO;
	lrHeater3_Analog: REAL;
	tspeed: REAL;
	TMR_ResetSafety: TON;
	tResetSafetyGuard: BOOL;
	TMR_StartupFan: TON;
	tElevatorUp: BOOL;
	tElevatorDown:BOOL;
	TMR_DelaySafetyModuleError: TON;
	Comm_OK: BOOL;
	TON_DelayAfterNetworkError: TON;
	REQ_RestartComm: BOOL;
	ReInitAllNodes: L_MC1P_ReinitAllNodes;
END_VAR
VAR
	Mach1_Drives_DB: Mach1_Drives;
	IDB_Dryer: Dryer;
	IDB_TrayFiller: TrayFiller;
END_VAR

NETWORK 0 LD TITLE: "DONE Network 1: Activating/deactivating MID-S/Trayfiller"
  LET g0 := TRUE;
  LET g1 := (g0 AND NOT Mach1_Safety.Status.Custom_ATF_Disabled);
  Mach1_AuxData.TrayfillerActive := g1;
  HMI_Var.TrayfillerActive := g1;
  Mach1_AuxData.MIDS_Active := (g0 AND TRUE);
END_NETWORK
NETWORK 1 LD TITLE: "DONE Network 2: Main Block FB100 TODO"
  LET i1 := fc_dinttotime(Mach1_Data.Timers.StartDelayAuxDrives,2);
  LET i2 := fc_dinttotime(Mach1_Data.Timers.StopDelayAuxDrives,2);
  tResetSafetyGuard := FB_Mach1(iStartResetSeparate := LST_General.AlwaysOff, iServiceButtonHasResetFunction := LST_General.AlwaysOff, iFirstCycle := LST_General.FirstCycle, iSignalPulse := LST_General.FF500ms, iAirPressureDoorsSeparate := LST_General.AlwaysOff, iEmergencyUnitOK := ((Mach1_AuxData.MIDS_Active AND Mach1_Safety.Status.EmergencyStopOK) OR NOT Mach1_AuxData.MIDS_Active), iDoorUnitOK := ((Mach1_AuxData.MIDS_Active AND Mach1_Safety.Status.DoorsOK) OR NOT Mach1_AuxData.MIDS_Active), iSTO_Enabled := Mach1_Safety.Status.STO_OK, iAirPressureOK := ((Mach1_AuxData.MIDS_Active AND LST_InputsOutputs.I100_0_AirpressureOK) OR NOT Mach1_AuxData.MIDS_Active), iSwitchService := Mach1_Safety.Status.ServiceMode, iButtonService := Mach1_Safety.Status.Service_ButtonAB, iStart1 := LST_InputsOutputs.I100_1_Pushbutton_start_OP0a, iStop1 := ((Mach1_AuxData.MIDS_Active AND LST_InputsOutputs.I100_2_Pushbutton_stop_OP0a) OR NOT Mach1_AuxData.MIDS_Active), iReset1 := LST_General.AlwaysOff, iAutoManual1 := LST_InputsOutputs.I100_3_Selector_switch_auto_manual_OP0a, iStart2 := (Mach1_AuxData.TrayfillerActive AND LST_InputsOutputs.I132_1_PB_Start_OP2a), iStop2 := (LST_InputsOutputs.I132_2_PB_Stop_OP2a OR NOT Mach1_AuxData.TrayfillerActive), iReset2 := LST_General.AlwaysOff, iAutoManual2 := LST_InputsOutputs.I132_3_SW_Auto_Man, iStart3 := LST_General.AlwaysOff, iStop3 := TRUE, iReset3 := LST_General.AlwaysOff, iAutoManual3 := LST_General.AlwaysOff, iPreDelayAfterEmergStop := T#4S, iPreStartDelayAuxDrives := i1, iPreStopDelayAuxDrives := i2, iPreDelayAfterSTOEnabled := T#2S, GenFlags := Mach1.GenFlags, oStart1 => LST_InputsOutputs.Q100_5_Signal_lamp_Start, oStop1 => LST_InputsOutputs.Q100_6_Signal_lamp_Stop, oCrossingDoorCircuit1 => tCrossDoorcircuit1, oStart2 => LST_InputsOutputs.Q132_0_SL_Start_OP2a, oStop2 => LST_InputsOutputs.Q132_1_SL_Stop_OP2a, oCrossingDoorCircuit2 => tCrossDoorcircuit2, oAlarm => tAlarmlamp);
END_NETWORK
NETWORK 2 LD
  LET g54 := TRUE;
  Mach1_Safety.Control.ResetSafetyGuard S= (g54 AND (mach1.Genflags.StartFlag OR tResetSafetyGuard));
  Mach1_Safety.Control.ResetSafetyGuard R= TMR_ResetSafety(IN := (g54 AND Mach1_Safety.Control.ResetSafetyGuard), PT := T#1S);
END_NETWORK
NETWORK 3 LD TITLE: "DONE Network 3 :Muting zones"
  LET g2 := (TRUE AND Mach1_AuxData.MainDriveHomed AND Mach1_AuxData.RollingDeviceHomed);
  Mach1_Safety.Control.Muting_zone1 := (g2 AND tCrossDoorcircuit1);
  Mach1_Safety.Control.Muting_zone2 := (g2 AND tCrossDoorcircuit1);
END_NETWORK
NETWORK 4 LD TITLE: "DONE NETWORK 4 (p1)Major alarms (start-up conditions)"
  Alarms_V5_1_100(Mach1_Alarms, (Mach1_AuxData.MIDS_Active AND NOT Mach1_Safety.Status.EmergencyStopOK), TRUE, Mach1_Alarms.Alm001, Mach1.GenFlags.MajorAlarm);
END_NETWORK
NETWORK 5 LD TITLE: "DONE NETWORK 4 (p2)Major alarms (start-up conditions)"
  Alarms_V5_1_100(Mach1_Alarms, (Mach1_AuxData.MIDS_Active AND Mach1_Safety.Status.EmergencyStopOK AND (NOT Mach1_Safety.Status.DoorsOK OR (Mach1_Safety.Status.ServiceMode AND NOT Mach1_AuxData.AllDrivesHomed AND NOT Mach1_Safety.Status.AllDoorsActuallyClosed))), TRUE, Mach1_Alarms.Alm002, Mach1.GenFlags.MinorAlarm);
END_NETWORK
NETWORK 6 LD TITLE: "DONE NETWORK 4 (p3)Major alarms (start-up conditions)"
  Alarms_V5_1_100(Mach1_Alarms, (Mach1_AuxData.MIDS_Active AND Mach1.Genflags.DelayAfterEmergStop AND NOT LST_InputsOutputs.I100_0_AirpressureOK), Mach1.GenFlags.StartFlag, Mach1_Alarms.Alm004, Mach1.GenFlags.MajorAlarm);
END_NETWORK
NETWORK 7 LD TITLE: "DONE NETWORK 4 (p4)Major alarms (start-up conditions)"
  Mach1_Safety.Control.ExternalRequestResetSafetyModule := (Alarms_V5_1_100(Mach1_Alarms, TMR_DelaySafetyModuleError(IN := (Mach1_AuxData.MIDS_Active AND (Mach1_Safety.Status.ErrorInInputModule OR Mach1_Safety.Status.ErrorInOutputModule)), PT := T#1S), TRUE, Mach1_Alarms.Alm009, Mach1.GenFlags.MinorAlarm) AND (FB_Mach1.iStart1 OR FB_Mach1.iStart2 OR FB_Mach1.iStart3));
END_NETWORK
NETWORK 8 LD
  Comm_OK := (Axis_MainDrive.xCommunicationOK AND Axis_SideCorrection.xCommunicationOK AND Axis_FeedFowardWrapper.xCommunicationOK AND Axis_OverrollingDevice.xCommunicationOK AND Axis_Bobbin.xCommunicationOK AND Axis_Fan.xCommunicationOK AND Axis_FeedForwardADS.xCommunicationOK AND Axis_FeedForwardATF.xCommunicationOK AND Axis_Elevator.xCommunicationOK);
END_NETWORK
NETWORK 9 LD TITLE: "DONE NETWORK 4 (p3)Major alarms (start-up conditions)"
  Alarms_V5_1_100(Mach1_Alarms, (LST_General.StartUpDelayPLC AND NOT Comm_OK), (Mach1.GenFlags.StartFlag OR NOT LST_General.StartUpDelayPLC OR Comm_OK), Mach1_Alarms.Alm011, Mach1.GenFlags.Warning);
END_NETWORK
NETWORK 10 LD
  LET g1 := TON_DelayAfterNetworkError(IN := (Mach1_Alarms.Alm011 AND NOT Mach1_Alarms.Alm011), PT := T#10000S);
  EtherCAT_Master.xRestart := g1;
  REQ_RestartComm S= g1;
END_NETWORK
NETWORK 11 LD
  ReInitAllNodes(xExecute := REQ_RestartComm, xInitCommunication := TRUE);
END_NETWORK
NETWORK 12 LD
  REQ_RestartComm R= (REQ_RestartComm AND Comm_OK);
END_NETWORK
NETWORK 13 LD TITLE: "TODO NETWORK 6"
  LET en1 := TRUE;
  IF en1 THEN MainDrive(); END_IF
  HMI_Var.Mach1.HourCounterRunning S= (en1 AND Mach1.GenFlags.DriveIsRunning);
END_NETWORK
NETWORK 14 LD TITLE: "DONE NETWORK 6: Drives"
  LET en1 := ;
  IF en1 THEN Mach1_Drives_DB(); END_IF
END_NETWORK
NETWORK 15 LD TITLE: "DONE NETWORK 7: Positioned stop leaf carrier"
  LET g3 := TRUE;
  Mach1_AuxData.MemStopLeafCarrier := (g3 AND HMI_Var.Btn_StopLeafCarrier AND ((Mach1.GenFlags.RunAuto AND Mach1.GenFlags.DriveIsRunning) OR Mach1_AuxData.MemStopLeafCarrier));
  tStopPositionLeafCarrier := (fc_CamC_CP_UDT(g3, HMI_Var.Mach1.Position, Mach1.GenFlags.Rotflag, Mach1_Data.CamControls.StopPostionLeafCarrier_CP) AND Mach1_Data.CamControls.StopPostionLeafCarrier_CP.Active AND Mach1_AuxData.MemStopLeafCarrier);
END_NETWORK
NETWORK 16 LD TITLE: "DONE NETWORK 8: Alarm Positioned stop leaf carrier"
  Mach1.GenFlags.StopDriveDirect S= Alarms_V5_1_100(Mach1_Alarms, tStopPositionLeafCarrier, NOT Mach1_AuxData.MemStopLeafCarrier, Mach1_Alarms.Alm054, Mach1.GenFlags.MinorAlarm);
END_NETWORK
NETWORK 17 LD TITLE: "DONE NETWORK 9: Positioned stop cleaning"
  LET g4 := TRUE;
  Mach1_AuxData.MemStopCleaning := (g4 AND HMI_Var.Btn_Cleaning AND ((Mach1.GenFlags.RunAuto AND Mach1.GenFlags.DriveIsRunning) OR Mach1_AuxData.MemStopCleaning));
  tStopPositionCleaning := (fc_CamC_CP_UDT(g4, HMI_Var.Mach1.Position, Mach1.GenFlags.Rotflag, Mach1_Data.CamControls.StopPostionCleaning_CP) AND Mach1_AuxData.MemStopCleaning);
END_NETWORK
NETWORK 18 LD TITLE: "DONE NETWORK 10: Alarm Positioned stop cleaning"
  Mach1.GenFlags.StopDriveDirect S= Alarms_V5_1_100(Mach1_Alarms, tStopPositionCleaning, NOT Mach1_AuxData.MemStopCleaning, Mach1_Alarms.Alm037, Mach1.GenFlags.MinorAlarm);
END_NETWORK
NETWORK 19 LD TITLE: "DONE NETWORK 11 (p1): Level bunch magazine alarms"
  LET en1 := ;
  IF en1 THEN ??? := Alarms_V5_1_100(Mach1_Alarms, Mach1_AuxData.IEC_TIMERS.TON_BunchLevelWarning(IN := (Mach1_AuxData.MIDS_Active AND Mach1.GenFlags.DelayAfterEmergStop AND NOT LST_InputsOutputs.I101_4_Level_bunch_magazine AND HMI_Var.Test_Prod AND NOT HMI_Var.Btn_Cleaning AND HMI_Var.Mach1.MuteNoBunchAlarm AND Mach1_Alarms.Alm036), PT := T#5S), (LST_InputsOutputs.I101_4_Level_bunch_magazine OR HMI_Var.Test_Prod OR HMI_Var.Btn_Cleaning OR HMI_Var.Mach1.MuteNoBunchAlarm OR Mach1_Alarms.Alm036), Mach1_Alarms.Alm073, Mach1.GenFlags.Warning); END_IF
END_NETWORK
NETWORK 20 LD TITLE: "DONE NETWORK 11 (p2): Level bunch magazine alarms"
  LET i1 := fc_dinttotime(Mach1_Data.Timers.BunchMagazineEmptyTime,0);
  Mach1.GenFlags.StopDriveDirect S= Alarms_V5_1_100(Mach1_Alarms, Mach1_AuxData.IEC_TIMERS.TON_BunchLevelAlarm(IN := (Mach1_AuxData.MIDS_Active AND Mach1.GenFlags.DelayAfterEmergStop AND NOT Mach1_Alarms.Alm036 AND NOT LST_InputsOutputs.I101_4_Level_bunch_magazine AND HMI_Var.Test_Prod AND NOT HMI_Var.Btn_Cleaning AND NOT HMI_Var.Mach1.MuteNoBunchAlarm), PT := i1), Mach1.GenFlags.StartFlag, Mach1_Alarms.Alm036, Mach1.GenFlags.MinorAlarm);
END_NETWORK
NETWORK 21 LD TITLE: "TODO NETWORK 12: SR Bunches (JL / rolling device / outfeed)"
  LET g119 := fc_camc_cp_udt(, HMI_Var.Mach1.Position, Mach1.GenFlags.Rotflag, Mach1_Data.CamControls.BunchDetection_CP);
  Mach1_AuxData.ShiftRegister.SR_bunch_present_position_3_outfeed R= (g119 AND Mach1_AuxData.ShiftRegister.SR_bunch_present_position_3_outfeed);
  LET g120 := (g119 AND Mach1_AuxData.ShiftRegister.SR_bunch_present_position_2_wrapping_device);
  Mach1_AuxData.ShiftRegister.SR_bunch_present_position_3_outfeed S= g120;
  Mach1_AuxData.ShiftRegister.SR_bunch_present_position_2_wrapping_device R= g120;
  LET g121 := (g119 AND Mach1_AuxData.ShiftRegister.SR_bunch_present_position_1_JL);
  Mach1_AuxData.ShiftRegister.SR_bunch_present_position_2_wrapping_device S= g121;
  Mach1_AuxData.ShiftRegister.SR_bunch_present_position_1_JL R= g121;
  Mach1_AuxData.ShiftRegister.SR_bunch_present_position_1_JL S= (g119 AND LST_InputsOutputs.I101_1_FC_Bunch_present);
  tBool := g119;
END_NETWORK
NETWORK 22 LD TITLE: "DONE NETWORK 13: Stop bunch infeed when cleaning is activated"
  HMI_Var.Btn_BunchSupply R= Mach1_AuxData.Edge.OSP_Emptying_Cleaning(CLK := HMI_Var.Btn_Cleaning);
END_NETWORK
NETWORK 23 LD TITLE: "DONE NETWORK 14: PNV Block bunch infeed"
  LET g5 := TRUE;
  LET g6 := (g5 AND TRUE);
  LET g7 := (fc_CamC_CP_UDT(g6, HMI_Var.Mach1.Position, LST_General.AlwaysOff, Mach1_Data.CamControls.BlockBunchInfeed_CP) AND TRUE);
  Mach1_AuxData.BlockBunchInfeed S= (g7 AND NOT HMI_Var.Btn_BunchSupply);
  Mach1_AuxData.BlockBunchInfeed R= (g7 AND HMI_Var.Btn_BunchSupply);
  Mach1_AuxData.BlockBunchInfeed S= (g6 AND NOT Mach1.GenFlags.DelayAfterEmergStop);
  PneumValveTerminalSMC.Pos2A := (g5 AND Mach1.GenFlags.EnablePneumEStop AND Mach1_AuxData.BlockBunchInfeed AND NOT Mach1_Alarms.Alm011);
END_NETWORK
NETWORK 24 LD TITLE: "DONE NETWORK 15: Muting of alarm ""No bunch"""
  LET i1 := INT_TO_WORD(Mach1_Data.Counters.BunchesFillBunchFeeder.SetValue);
  Mach1_AuxData.NumberOfMutingCyclesReached := Mach1_AuxData.COUNTERS.RepetitionMuteNuBunch(CD := (ATD_SR(Mach1_Alarms.Alm041, (tBool AND (NOT HMI_Var.Test_Prod OR HMI_Var.Btn_Cleaning OR Mach1_AuxData.ShiftRegister.SR_bunch_present_position_1_JL OR NOT HMI_Var.Btn_BunchSupply OR Mach1_AuxData.NumberOfMutingCyclesReached)), hmi_var.mach1.MuteNoBunchAlarm) AND tBool AND HMI_Var.Test_Prod AND NOT HMI_Var.Btn_Cleaning AND NOT Mach1_AuxData.ShiftRegister.SR_bunch_present_position_1_JL), LOAD := Mach1_Alarms.Alm041, PV := i1);
END_NETWORK
NETWORK 25 LD TITLE: "DONE NETWORK 16 (p1): Alarms Bunch"
  LET i1 := INT_TO_WORD(Mach1_Data.Counters.MaxRepetitionNoBunch.SetValue);
  Mach1.GenFlags.StopDriveDirect S= Alarms_V5_1_100(Mach1_Alarms, ((Mach1_AuxData.COUNTERS.RepetitionNoBunch(CD := (tBool AND HMI_Var.Test_Prod AND NOT HMI_Var.Btn_Cleaning AND NOT HMI_Var.Mach1.MuteNoBunchAlarm AND NOT Mach1_AuxData.ShiftRegister.SR_bunch_present_position_1_JL), LOAD := ((tBool AND (NOT HMI_Var.Test_Prod OR HMI_Var.Btn_Cleaning OR Mach1_AuxData.ShiftRegister.SR_bunch_present_position_1_JL OR NOT HMI_Var.Btn_BunchSupply OR hmi_var.mach1.MuteNoBunchAlarm)) OR (Mach1.GenFlags.StartFlag AND Mach1_Alarms.Alm041)), PV := i1) AND Mach1_AuxData.AllDrivesHomed) AND NOT HMI_Var.Mach1.MuteNoBunchAlarm), Mach1.GenFlags.StartFlag, Mach1_Alarms.Alm041, Mach1.GenFlags.MinorAlarm);
END_NETWORK
NETWORK 26 LD TITLE: "DONE NETWORK 16 (p2): Alarms Bunch"
  Mach1.GenFlags.StopDriveDirect S= Alarms_V5_1_100(Mach1_Alarms, (tBool AND NOT Mach1_AuxData.PhotocellBunchHasBeenOff AND HMI_Var.Btn_BunchSupply AND Mach1_AuxData.AllDrivesHomed), Mach1.GenFlags.StartFlag, Mach1_Alarms.Alm042, Mach1.GenFlags.MinorAlarm);
END_NETWORK
NETWORK 27 LD TITLE: "DONE NETWORK 16 (p3): Alarms Bunch"
  ATD_SR(NOT LST_InputsOutputs.I101_1_FC_Bunch_present, tBool, Mach1_AuxData.PhotocellBunchHasBeenOff);
END_NETWORK
NETWORK 28 LD
END_NETWORK
NETWORK 29 LD TITLE: "DONE NETWORK 17 (p1): Alarms: Cigar fault"
  LET i1 := INT_TO_WORD(Mach1_Data.Counters.MaxRepetitionNoCigars.SetValue);
  Mach1.GenFlags.StopDriveDirect S= Alarms_V5_1_100(Mach1_Alarms, (Mach1_AuxData.COUNTERS.RepetitionNoCigar(CD := (fc_CamC_CP_UDT(, HMI_Var.Mach1.Position, Mach1.GenFlags.Rotflag, Mach1_Data.CamControls.CigarDetection_CP) AND HMI_Var.Test_Prod AND NOT HMI_Var.Btn_Cleaning AND Mach1_AuxData.ShiftRegister.SR_bunch_present_position_3_outfeed AND NOT LST_InputsOutputs.I101_2_Cigar_present), LOAD := ((tBool AND (NOT HMI_Var.Test_Prod OR HMI_Var.Btn_Cleaning OR (Mach1_AuxData.ShiftRegister.SR_bunch_present_position_3_outfeed AND LST_InputsOutputs.I101_2_Cigar_present))) OR (Mach1.GenFlags.StartFlag AND Mach1_Alarms.Alm046)), PV := i1) AND Mach1_AuxData.AllDrivesHomed), Mach1.GenFlags.StartFlag, Mach1_Alarms.Alm046, Mach1.GenFlags.MinorAlarm);
END_NETWORK
NETWORK 30 LD TITLE: "DONE NETWORK 17 (p2): Alarms: Cigar fault"
  Mach1.GenFlags.StopDriveDirect S= Alarms_V5_1_100(Mach1_Alarms, (tbool AND NOT Mach1_AuxData.PhotocellCigarHasBeenOff AND Mach1_AuxData.AllDrivesHomed), Mach1.GenFlags.StartFlag, Mach1_Alarms.Alm047, Mach1.GenFlags.MinorAlarm);
END_NETWORK
NETWORK 31 LD TITLE: "DONE NETWORK 17 (p3): Alarms: Cigar fault"
  ATD_SR(NOT LST_InputsOutputs.I101_2_Cigar_present, tbool, Mach1_AuxData.PhotocellCigarHasBeenOff);
END_NETWORK
NETWORK 32 LD TITLE: "DONE NETWORK 18: Production counter"
  HMI_Var.Mach1.PRDCounterIncr S= (tBool AND Mach1_AuxData.ShiftRegister.SR_bunch_present_position_3_outfeed AND LST_InputsOutputs.I101_2_Cigar_present);
END_NETWORK
NETWORK 33 LD TITLE: "DONE NETWORK 19 (p1): Set cigar present in checkRegister"
  LET g124 := TRUE;
  db_CheckRegister.Positie[1].Infeed.Cigar_present_infeed S= (g124 AND tCampulseCigarPresent AND LST_InputsOutputs.I101_2_Cigar_present);
  Mach1_AuxData.MemCigarAtCrossOver S= (g124 AND LST_InputsOutputs.I133_2_Cigar_detected_at_cross_over);
  LET g125 := Mach1_AuxData.Edge.OSP_DryerZeroPoint(CLK := (g124 AND LST_InputsOutputs.I133_1_PROX_zero_position_transport_ADS));
  LET g126 := (g125 AND Mach1_AuxData.MemCigarAtCrossOver);
  db_CheckRegister.Positie[CTE.posCigarPresentOutfeed].Outfeed.Cigar_present_outfeed S= g126;
  Mach1_AuxData.MemCigarAtCrossOver R= g126;
  Mach1_AuxData.PreviousCycleHasOutfeedError R= g125;
  Mach1_AuxData.PreviousCycleHasOutfeedError S= (g125 AND Mach1_AuxData.CurrentCycleHasOutfeedError);
  LET en1 := g125;
  IF en1 THEN fc_CheckRegister(); END_IF
  Mach1_AuxData.CurrentCycleHasOutfeedError R= g125;
  Mach1_AuxData.CurrentCycleHasOutfeedError S= (g125 AND db_CheckRegister.CheckRegisterError);
END_NETWORK
NETWORK 34 LD TITLE: "DONE NETWORK 20: Start Fan"
  LET g109 := (Mach1.GenFlags.EnableAuxDrive AND HMI_Var.Test_Prod AND NOT HMI_Var.Btn_Cleaning);
  Mach1_Data.Drives.Fan.Control.StartAuto := g109;
  TMR_StartupFan(IN := g109, PT := T#5S);
END_NETWORK
NETWORK 35 LD
  mach1.Genflags.StopDriveDirect S= Alarms_V5_1_100(Mach1_Alarms, (NOT HMI_Var.Btn_Cleaning AND Mach1.GenFlags.EnableAuxDrive AND HMI_Var.Test_Prod AND NOT TMR_StartupFan.Q), TRUE, Mach1_Alarms.Alm034, mach1.Genflags.MinorAlarm);
END_NETWORK
NETWORK 36 LD TITLE: "DONE NETWORK 21: Blocking glue rod"
  LET g12 := (Mach1.GenFlags.EnablePneumEStop AND Mach1_Safety.Status.DoorsOK);
  PneumValveTerminalSMC.Pos3A := (g12 AND (NOT Mach1_AuxData.ShiftRegister.SR_bunch_present_position_2_wrapping_device OR NOT HMI_Var.Test_Prod OR HMI_Var.Btn_Cleaning) AND Mach1_AuxData.AllDrivesHomed AND NOT Mach1_Alarms.Alm011);
  PneumValveTerminalSMC.Pos3B := (g12 AND NOT PneumValveTerminalSMC.Pos3A);
END_NETWORK
NETWORK 37 LD TITLE: "DONE NETWORK 22 (p1): Insert needle"
  PneumValveTerminalSMC.Pos4A := (fc_CamC_LS_UDT((Mach1_Safety.Status.DoorsOK AND Mach1.GenFlags.EnablePneumEStop), HMI_Var.Mach1.ActualSpeed, HMI_Var.Mach1.Position, Mach1.GenFlags.Rotflag, Mach1_Data.CamControls.InserNeedle_CLS) AND Mach1_AuxData.AllDrivesHomed AND NOT Mach1_Alarms.Alm011);
END_NETWORK
NETWORK 38 LD TITLE: "DONE NETWORK 22 (p2): Insert needle"
  PneumValveTerminalSMC.Pos4B := (Mach1_Safety.Status.DoorsOK AND Mach1.GenFlags.EnablePneumEStop AND NOT PneumValveTerminalSMC.Pos4A);
END_NETWORK
NETWORK 39 LD TITLE: "DONE NETWORK 23 (p1): Bunch positioner"
  PneumValveTerminalSMC.Pos5A := (fc_CamC_LS_UDT((Mach1_Safety.Status.DoorsOK AND Mach1.GenFlags.EnablePneumEStop), HMI_Var.Mach1.ActualSpeed, HMI_Var.Mach1.Position, Mach1.GenFlags.Rotflag, Mach1_Data.CamControls.BunchPositioner_CLS) AND Mach1_AuxData.AllDrivesHomed AND NOT Mach1_Alarms.Alm011);
END_NETWORK
NETWORK 40 LD TITLE: "DONE NETWORK 23 (p2): Bunch positioner"
  PneumValveTerminalSMC.Pos5B := (Mach1_Safety.Status.DoorsOK AND Mach1.GenFlags.EnablePneumEStop AND NOT PneumValveTerminalSMC.Pos5A);
END_NETWORK
NETWORK 41 LD TITLE: "DONE NETWORK 24: Manual glue pumping"
  LET g103 := Mach1_AuxData.EnableGlueSprayCalibration;
  LET g104 := (g103 AND TRUE AND (HMI_Var.Mach1.GlueStart OR HMI_Var.Mach1.GlueStop OR HMI_Var.Mach1.GlueReset OR HMI_Var.Mach1.SprayStart OR HMI_Var.Mach1.SprayStop OR HMI_Var.Mach1.SprayReset OR Mach1_AuxData.ScreenForOperatorSettingsActivated));
  Mach1_AuxData.ScreenForOperatorSettingsActivated := g104;
  Mach1.GenFlags.StopDriveDirect S= g104;
  LET en1 := (g103 AND (HMI_Var.Mach1.GlueReset OR NOT LST_InputsOutputs.I100_2_Pushbutton_stop_OP0a));
  IF en1 THEN Mach1_Data.Settings.Ints.ActualNumberOfGluePulses := MOVE(0); END_IF
  LET en2 := (g103 AND Mach1.GenFlags.EnablePneumEStop AND (((HMI_Var.Mach1.GlueStart OR LST_InputsOutputs.I100_4_Pushbutton_request_glue_OP0a) AND NOT LST_General.FF500ms) OR Mach1_AuxData.GlueWeighingCycleStarted) AND NOT HMI_Var.Mach1.GlueStop AND NOT HMI_Var.Mach1.GlueReset AND LST_InputsOutputs.I100_2_Pushbutton_stop_OP0a);
  IF en2 THEN Mach1_AuxData.GlueWeighingCycleStarted := (Mach1_Data.Settings.Ints.ActualNumberOfGluePulses < Mach1_Data.Settings.Ints.MaxNumberOfGluePulses); END_IF
  LET en3 := (Mach1_AuxData.Edge.OSN_Gluepump(CLK := (g103 AND PneumValveTerminalSMC.Pos6A)) AND Mach1_AuxData.GlueWeighingCycleStarted);
  IF en3 THEN Mach1_Data.Settings.Ints.ActualNumberOfGluePulses := (Mach1_Data.Settings.Ints.ActualNumberOfGluePulses + 1); END_IF
END_NETWORK
NETWORK 42 LD TITLE: "DONE NETWORK 25: Continuous Glueing"
  LET g15 := TRUE;
  LET g16 := (NOT(Mach1_AuxData.Edge.OSPushbuttonGlue(CLK := (g15 AND (LST_InputsOutputs.I100_4_Pushbutton_request_glue_OP0a OR Mach1_AuxData.IEC_TIMERS.TON_StopContGluePumping.Q)))) AND Mach1.GenFlags.EnablePneumEStop AND NOT Mach1.GenFlags.DriveIsRunning AND NOT Mach1_AuxData.ScreenForOperatorSettingsActivated AND (LST_InputsOutputs.I100_4_Pushbutton_request_glue_OP0a OR Mach1_AuxData.IEC_TIMERS.DelayContiniousGluePumping.Q));
  Mach1_AuxData.MemContinuousGluePumping := g16;
  Mach1_AuxData.IEC_TIMERS.DelayContiniousGluePumping(IN := g16, PT := T#3S);
  Mach1_AuxData.IEC_TIMERS.TON_StopContGluePumping(IN := (g15 AND Mach1_AuxData.MemContinuousGluePumping), PT := T#120S);
END_NETWORK
NETWORK 43 LD TITLE: "DONE NETWORK 26: PNV Glue pump 1+2+3"
  LET g1 := (((fc_CamC_CC_UDT(Mach1.GenFlags.EnablePneumEStop, HMI_Var.Mach1.Position, Mach1_Data.CamControls.GluePump123_C) AND Mach1_AuxData.ShiftRegister.SR_bunch_present_position_1_JL AND HMI_Var.Test_Prod AND NOT HMI_Var.Btn_Cleaning AND NOT Mach1_AuxData.MemContinuousGluePumping AND NOT Mach1_AuxData.ScreenForOperatorSettingsActivated) OR (Mach1.GenFlags.EnablePneumEStop AND ((LST_General.FF500ms AND Mach1_AuxData.MemContinuousGluePumping) OR (LST_General.FF500ms AND Mach1_AuxData.GlueWeighingCycleStarted)))) AND NOT Mach1_Alarms.Alm011);
  PneumValveTerminalSMC.Pos6A := g1;
  LST_InputsOutputs.Q101_2_Enable_GluePump := g1;
END_NETWORK
NETWORK 44 LD TITLE: "DONE NETWORK 27: PNV Glue pump 4"
  PneumValveTerminalSMC.Pos10A := (((fc_CamC_CC_UDT(Mach1.GenFlags.EnablePneumEStop, HMI_Var.Mach1.Position, Mach1_Data.CamControls.GluePump4_C) AND Mach1_AuxData.ShiftRegister.SR_bunch_present_position_1_JL AND HMI_Var.Test_Prod AND NOT HMI_Var.Btn_Cleaning AND NOT Mach1_AuxData.MemContinuousGluePumping AND NOT Mach1_AuxData.ScreenForOperatorSettingsActivated) OR (Mach1.GenFlags.EnablePneumEStop AND ((LST_General.FF500ms AND Mach1_AuxData.MemContinuousGluePumping) OR (LST_General.FF500ms AND Mach1_AuxData.GlueWeighingCycleStarted)))) AND NOT Mach1_Alarms.Alm011);
END_NETWORK
NETWORK 45 LD TITLE: "DONE NETWORK 28: PNV Glue pump 5"
  PneumValveTerminalSMC.Pos11A := (((fc_CamC_CC_UDT(Mach1.GenFlags.EnablePneumEStop, HMI_Var.Mach1.Position, Mach1_Data.CamControls.GluePump5_C) AND Mach1_AuxData.ShiftRegister.SR_bunch_present_position_1_JL AND HMI_Var.Test_Prod AND NOT HMI_Var.Btn_Cleaning AND NOT Mach1_AuxData.MemContinuousGluePumping AND NOT Mach1_AuxData.ScreenForOperatorSettingsActivated) OR (Mach1.GenFlags.EnablePneumEStop AND ((LST_General.FF500ms AND Mach1_AuxData.MemContinuousGluePumping) OR (LST_General.FF500ms AND Mach1_AuxData.GlueWeighingCycleStarted)))) AND NOT Mach1_Alarms.Alm011);
END_NETWORK
NETWORK 46 LD TITLE: "DONE NETWORK 29: PNV Small gripper"
  PneumValveTerminalSMC.Pos7A := (fc_CamC_LS_UDT(Mach1.GenFlags.EnablePneumEStop, HMI_Var.Mach1.ActualSpeed, HMI_Var.Mach1.Position, Mach1.GenFlags.Rotflag, Mach1_Data.CamControls.SmallGripper_CLS) AND Mach1_AuxData.AllDrivesHomed AND NOT Mach1_Alarms.Alm011);
END_NETWORK
NETWORK 47 LD TITLE: "DONE NETWORK 30: Big gripper"
  PneumValveTerminalSMC.Pos8A := (fc_CamC_LS_UDT(Mach1.GenFlags.EnablePneumEStop, HMI_Var.Mach1.ActualSpeed, HMI_Var.Mach1.Position, Mach1.GenFlags.Rotflag, Mach1_Data.CamControls.BigGripper_CLS) AND Mach1_AuxData.AllDrivesHomed AND NOT Mach1_Alarms.Alm011);
END_NETWORK
NETWORK 48 LD TITLE: "TODO NETWORK 31: Blow off wrapper"
  PneumValveTerminalSMC.Pos9A := (fc_CamC_CC_UDT(Mach1.GenFlags.EnablePneumEStop, HMI_Var.Mach1.Position, Mach1_Data.CamControls.BlowOffWrapper_C) AND NOT Mach1_Alarms.Alm011);
END_NETWORK
NETWORK 49 LD TITLE: "DONE NETWORK 32: Blow off bobbin"
  PneumValveTerminalSMC.Pos1A := (fc_CamC_CC_UDT((Mach1.GenFlags.EnablePneumEStop AND Mach1.GenFlags.DriveIsRunning), HMI_Var.Mach1.Position, Mach1_Data.CamControls.BlowOffBobine_C) AND NOT Mach1_Alarms.Alm011);
END_NETWORK
NETWORK 50 LD TITLE: "DONE NETWORK 33:"
  LET en1 := ;
  IF en1 THEN AHWF(); END_IF
END_NETWORK
NETWORK 51 LD TITLE: "TODO NETWORK 34: OBSOLETE"
END_NETWORK
NETWORK 52 LD TITLE: "DONE NETWORK 35: Main FB:  Dryer-trayfiller"
  LET en1 := ;
  IF en1 THEN (Mach1_AuxData.COUNTERS.EmptyingCycles.CV < 105); END_IF
  LET g105 := IDB_Dryer(iGenFlags := Mach1.GenFlags, iMachineStarted := (Mach1.GenFlags.EnableAuxDrive AND Mach1_Safety.Status.DoorsOK AND NOT Mach1.GenFlags.StopFlag), iSwitchDryer := HMI_Var.Btn_DryerOn, iDryerClosed := LST_InputsOutputs.I133_0_PROX_Dryer_closed, iStartFeedForward := fc_CamC_CP_UDT(, HMI_Var.Mach1.Position, Mach1.GenFlags.Rotflag, Mach1_Data.CamControls.FeedforwardDryer_CP), iStopFeedForward := (((NOT Mach1.GenFlags.EnableAuxDrive OR en1 OR NOT Trayfiller_Data.commInterface.Permission OR NOT Mach1_Safety.Status.DoorsOK) AND LST_InputsOutputs.I133_1_PROX_zero_position_transport_ADS) OR Mach1_Alarms.Alm048), iPermissionDownstream := (Trayfiller_Data.commInterface.Permission AND NOT Mach1_Alarms.Alm053), iSetPowerHeater1 := Mach1_Data.Dryer.Heater1.SetHeaterPower, iSetPowerHeater2 := Mach1_Data.Dryer.Heater2.SetHeaterPower, iSetPowerHeater3 := Mach1_Data.Dryer.Heater3.SetHeaterPower, iPowerOrAnalog := TRUE, iSpeedForEmptying := 100, oEnableHeaters => HMI_Var.Mach1.HeatersActive, oPowerHeater1 => tHeater1Word, oPowerHeater2 => tHeater2Word, oPowerHeater3 => tHeater3Word);
  LST_InputsOutputs.Q132_2_Enable_power_controllers := (g105 AND HMI_Var.Mach1.HeatersActive);
  LET en2 := g105;
  IF en2 THEN (Mach1_Data.Dryer.Heater1.SetHeaterPower >= 350); END_IF
  LET en3 := en2;
  IF en3 THEN Mach1_Data.Dryer.Heater1.SetHeaterPower := MOVE(350); END_IF
  LET en4 := g105;
  IF en4 THEN (Mach1_Data.Dryer.Heater2.SetHeaterPower >= 350); END_IF
  LET en5 := en4;
  IF en5 THEN Mach1_Data.Dryer.Heater2.SetHeaterPower := MOVE(350); END_IF
  LET en6 := g105;
  IF en6 THEN (Mach1_Data.Dryer.Heater3.SetHeaterPower >= 350); END_IF
  LET en7 := en6;
  IF en7 THEN Mach1_Data.Dryer.Heater3.SetHeaterPower := MOVE(350); END_IF
END_NETWORK
NETWORK 53 LD TITLE: "DONE NETWORK 36: CT Fan dryer"
  LST_InputsOutputs.Q132_4_CT_Fan_dryer := (Mach1_AuxData.TrayfillerActive AND Mach1.GenFlags.EnableAuxDrive AND HMI_Var.Btn_DryerOn);
END_NETWORK
NETWORK 54 LD TITLE: "TODO NETWORK 37:"
  // dryer speed: 100rpm ->1000 0.1rpm
  // max AO-value: 2^14=16384
  LET g40 := TRUE;
  LET i1 := DINT_TO_REAL(HMI_Var.Mach1.ActualSpeedDryer);
  LET en1 := g40;
  IF en1 THEN DRYER_Scaling_Speed(IN := i1, IN_MIN := 0, IN_MAX := 1000, OUT_MIN := 0, OUT_MAX := 1, OUT => lrDryer_ScaledSpeed); END_IF
  LET en2 := g40;
  IF en2 THEN DRYER_SCALING_Heater1(IN := tHeater1Word, IN_MIN := 0, IN_MAX := 1500, OUT_MIN := 0, OUT_MAX := 1, OUT => lrHeater1_ScaledPower); END_IF
  LET i2 := REAL_TO_INT(lrHeater1_ScaledPower*lrDryer_ScaledSpeed*1500);
  LET en3 := en2;
  IF en3 THEN HMI_Var.Mach1.ActHeater1 := MOVE(i2); END_IF
  LET en4 := en3;
  IF en4 THEN DRYER_SCALING_Heater1_Analog(IN := lrDryer_ScaledSpeed*lrHeater1_ScaledPower*1500, IN_MIN := 0, IN_MAX := 1500, OUT_MIN := 0, OUT_MAX := 16384, OUT => lrHeater1_Analog); END_IF
  LET i3 := REAL_TO_WORD(lrHeater1_Analog);
  LET en5 := en4;
  IF en5 THEN %QW105 := MOVE(i3); END_IF
  LET en6 := g40;
  IF en6 THEN DRYER_SCALING_Heater2(IN := tHeater2Word, IN_MIN := 0, IN_MAX := 1500, OUT_MIN := 0, OUT_MAX := 1, OUT => lrHeater2_ScaledPower); END_IF
  LET i4 := REAL_TO_INT(lrHeater2_ScaledPower*lrDryer_ScaledSpeed*1500);
  LET en7 := en6;
  IF en7 THEN HMI_Var.Mach1.ActHeater2 := MOVE(i4); END_IF
  LET en8 := en7;
  IF en8 THEN DRYER_SCALING_Heater2_Analog(IN := lrDryer_ScaledSpeed*lrHeater2_ScaledPower*1500, IN_MIN := 0, IN_MAX := 1500, OUT_MIN := 0, OUT_MAX := 16384, OUT => lrHeater2_Analog); END_IF
  LET i5 := REAL_TO_WORD(lrHeater2_Analog);
  LET en9 := en8;
  IF en9 THEN %QW106 := MOVE(i5); END_IF
  LET en10 := g40;
  IF en10 THEN DRYER_SCALING_Heater3(IN := tHeater3Word, IN_MIN := 0, IN_MAX := 1500, OUT_MIN := 0, OUT_MAX := 1, OUT => lrHeater3_ScaledPower); END_IF
  LET i6 := REAL_TO_INT(lrHeater3_ScaledPower*lrDryer_ScaledSpeed*1500);
  LET en11 := en10;
  IF en11 THEN HMI_Var.Mach1.ActHeater3 := MOVE(i6); END_IF
  LET en12 := en11;
  IF en12 THEN DRYER_SCALING_Heater2_Analog(IN := lrDryer_ScaledSpeed*lrHeater3_ScaledPower*1500, IN_MIN := 0, IN_MAX := 1500, OUT_MIN := 0, OUT_MAX := 16384, OUT => lrHeater3_Analog); END_IF
  LET i7 := REAL_TO_WORD(lrHeater3_Analog);
  LET en13 := en12;
  IF en13 THEN %QW107 := MOVE(i7); END_IF
END_NETWORK
NETWORK 55 LD TITLE: "DONE NETWORK 38 (p1): Alarms dryer"
  LET en1 := (Mach1.GenFlags.EnableAuxDrive AND NOT Mach1_Alarms.Alm048 AND ((Mach1.Genflags.DelayAfterSTO AND IDB_Dryer.oFeedForward) OR mach1.Genflags.DriveIsRunning) AND NOT LST_InputsOutputs.I133_1_PROX_zero_position_transport_ADS);
  IF en1 THEN (Mach1_Data.Drives.FeedForwardADS.Control.AutoSpeed >= 10); END_IF
  Mach1.GenFlags.StopDriveDirect S= RuntimeGuard_V5_1_100(Mach1_Alarms, (Mach1_AuxData.TrayfillerActive AND ((IDB_Dryer.oFeedForward AND Mach1.Genflags.DelayAfterSTO) OR mach1.Genflags.DriveIsRunning) AND (Mach1_AuxData.AllDrivesHomed OR NOT Mach1_AuxData.MIDS_Active)), LST_General.AlwaysOff, en1, T#10S, Mach1.GenFlags.StartFlag, Mach1_Alarms.Alm048, Mach1.GenFlags.MinorAlarm, Mach1_AuxData.IEC_TIMERS.RuntimeGuardFeedforwardDryer, oForwardUnguarded => tBool, oForwardGuarded => Mach1_Data.Drives.FeedForwardADS.Control.StartAuto, oReverseUnguarded => tBool, oReverseGuarded => tBool);
END_NETWORK
NETWORK 56 LD TITLE: "DONE NETWORK 38 (p2): Alarms dryer"
  Mach1.GenFlags.StopDriveDirect S= (Alarms_V5_1_100(Mach1_Alarms, (Mach1_AuxData.TrayfillerActive AND Mach1.GenFlags.DelayAfterEmergStop AND IDB_Dryer.oFaultDryerOpened), TRUE, Mach1_Alarms.Alm049, Mach1.GenFlags.MinorAlarm) AND Mach1_AuxData.AllDrivesHomed);
END_NETWORK
NETWORK 57 LD TITLE: "TODO NETWORK 38 (p3): Alarms dryer"
  LET en1 := (mach1.Genflags.DelayAfterEmergStop AND HMI_Var.Test_Prod AND Mach1_AuxData.TrayfillerActive);
  IF en1 THEN (Mach1_Data.Counters.MaxRepetitionNoCigarsDryer.SetValue > 0); END_IF
  LET g123 := Alarms_V5_1_100(Mach1_Alarms, (en1 AND db_CheckRegister.CheckRegisterError AND NOT Mach1_AuxData.PreviousCycleHasOutfeedError), Mach1.GenFlags.StartFlag, Mach1_Alarms.Alm053, Mach1.GenFlags.MinorAlarm);
  Mach1.GenFlags.StopDriveDirect S= g123;
  db_CheckRegister.CheckRegisterError R= g123;
END_NETWORK
NETWORK 58 LD TITLE: "DONE NETWORK 38 (p4): Alarms dryer"
  Mach1.GenFlags.StopDriveDirect S= Alarms_V5_1_100(Mach1_Alarms, Mach1_AuxData.IEC_TIMERS.TON_DryerSwitchedOff(IN := (Mach1_AuxData.TrayfillerActive AND HMI_Var.Test_Prod AND NOT HMI_Var.Btn_DryerOn), PT := T#5S), Mach1.GenFlags.StartFlag, Mach1_Alarms.Alm058, Mach1.GenFlags.MinorAlarm);
END_NETWORK
NETWORK 59 LD TITLE: "TODO NETWORK 39: Analog setpoint feedforward dryer"
  LET en1 := ;
  IF en1 THEN ??? := SpeedCalculationDryer(); END_IF
END_NETWORK
NETWORK 60 LD TITLE: "TODO NETWORK 40: Analog setpoint feedforward trayfiller"
  LET en1 := ;
  IF en1 THEN ??? := SpeedCalculationTrayfiller(); END_IF
END_NETWORK
NETWORK 61 LD TITLE: "DONE NETWORK 41: Empty trayfiller"
  HMI_Var.Btn_Cleaning R= Mach1_AuxData.COUNTERS.EmptyingCycles(CD := (HMI_Var.Btn_Cleaning AND LST_InputsOutputs.I133_1_PROX_zero_position_transport_ADS), LOAD := NOT HMI_Var.Btn_Cleaning, PV := 194);
END_NETWORK
NETWORK 62 LD TITLE: "DONE NETWORK 42: Main block Trayfiller"
  LET en1 := ;
  IF en1 THEN (Mach1_AuxData.COUNTERS.EmptyingCycles.CV < 106); END_IF
  LET en2 := ;
  IF en2 THEN (Mach1_AuxData.COUNTERS.EmptyingCycles.CV < 106); END_IF
  IDB_TrayFiller(iGenFlags := Mach1.GenFlags, iMachineStarted := (Mach1.GenFlags.EnableAuxDrive AND NOT Mach1.GenFlags.StopFlag), iButtonChangeTray := LST_General.AlwaysOff, iButtonTrayDown := LST_InputsOutputs.I132_6_Tray_down, iButtonTrayUp := LST_InputsOutputs.I132_7_Tray_up, iCigarAtCrossover := (LST_InputsOutputs.I133_2_Cigar_detected_at_cross_over OR en1), iStartFeedForward := ((LST_InputsOutputs.I133_1_PROX_zero_position_transport_ADS OR en2) AND Mach1_Safety.Status.DoorsOK), iStopFeedForward := LST_InputsOutputs.I133_3_PROX_zero_position_transport_ATF, iCigarAtInpusher := LST_InputsOutputs.I133_4_Cigar_detected_at_inpusher, iRpsInpusher := LST_InputsOutputs.I133_6_PROX_inpusher_retracted, iEpsInpusher := LST_InputsOutputs.I133_7_PROX_inpusher_at_tray, iGuardInpusher := TRUE, iPsElevatorUp := LST_InputsOutputs.I136_0_PROX_Elevator_above, iPsElevatorDown := LST_InputsOutputs.I136_1_PROX_Elevator_below, iPulseCounterElevator := LST_InputsOutputs.I136_2_PROX_pulse_counter_elevator, iFcGuardTrayOnElev := LST_InputsOutputs.I136_3_FC_Position_tray_OK, iRowHeight := Mach1_Data.TrayFiller.RowHeight, iSetNumberOfRows := Mach1_Data.Trayfiller.SetNumberOfRows, iInitialDescentValue := Mach1_Data.Trayfiller.InitialDescentValue, iLightCurtainInpusher := Mach1_Safety.Status.Door_switch17, iLightCurtainElevator := Mach1_Safety.Status.Door_switch18, iPsInfeedConvAtInit := LST_InputsOutputs.I136_4_PROX_Infeed_conveyor_initial_position, iPsInfeedConvAtElev := LST_InputsOutputs.I136_5_PROX_Infeed_conveyor_at_elevator, iFcGuardTrayFromElev := LST_InputsOutputs.I136_6_FC_Guard_tray_from_elevator, iFcOutfeedConvFull := LST_InputsOutputs.I136_7_FC_Outfeed_conveyor_full, iTestProd := TRUE, ioActNumberOfRows := HMI_Var.Mach1.ActNumberOfRows, oValveTiltInpusher => LST_InputsOutputs.Q132_7_PNV_tilting_inpusher);
END_NETWORK
NETWORK 63 LD
  Mach1_Data.Drives.FeedForwardATF.Control.StartAuto := IDB_TrayFiller.oFeedForwardMotor;
END_NETWORK
NETWORK 64 LD TITLE: "DONE NETWORK 43: Selection of inpusher runtimeguard time"
  LET g20 := IDB_TrayFiller.oValveInpusher;
  LET en1 := g20;
  IF en1 THEN tTime1 := MOVE(T#1S); END_IF
  LET en2 := NOT(g20);
  IF en2 THEN tTime1 := MOVE(T#5S); END_IF
END_NETWORK
NETWORK 65 LD TITLE: "DONE NETWORK 44 (p1): Runtimeguard trayfiller"
  Mach1.GenFlags.StopDriveDirect S= RuntimeGuard_V5_1_100(Mach1_Alarms, (Mach1_AuxData.TrayfillerActive AND IDB_TrayFiller.oValveInpusher AND Mach1_AuxData.AllDrivesHomed), (Mach1_AuxData.TrayfillerActive AND NOT IDB_TrayFiller.oValveInpusher AND Mach1_AuxData.AllDrivesHomed), (Mach1_AuxData.TrayfillerActive AND Mach1.GenFlags.EnablePneumEStop AND ((IDB_TrayFiller.oValveInpusher AND NOT LST_InputsOutputs.I133_7_PROX_inpusher_at_tray) OR (NOT IDB_TrayFiller.oValveInpusher AND NOT LST_InputsOutputs.I133_6_PROX_inpusher_retracted))), T#3S, Mach1.GenFlags.StartFlag, Mach1_Alarms.Alm050, Mach1.GenFlags.MinorAlarm, Mach1_AuxData.IEC_TIMERS.RuntimeguardInpusher, oForwardUnguarded => LST_InputsOutputs.Q132_6_PNV_Inpusher, oReverseUnguarded => tBool, oReverseGuarded => tBool);
END_NETWORK
NETWORK 66 LD TITLE: "DONE NETWORK 44 (p2): Runtimeguard trayfiller"
  Mach1.GenFlags.StopDriveDirect S= RuntimeGuard_V5_1_100(Mach1_Alarms, (Mach1_AuxData.TrayfillerActive AND IDB_TrayFiller.oElevatorMotorUp AND Mach1_AuxData.AllDrivesHomed), (Mach1_AuxData.TrayfillerActive AND IDB_TrayFiller.oElevatorMotorDown AND Mach1_AuxData.AllDrivesHomed), TRUE, T#15S, Mach1.GenFlags.StartFlag, Mach1_Alarms.Alm052, Mach1.GenFlags.MinorAlarm, Mach1_AuxData.IEC_TIMERS.RuntimeGuardElevator, oForwardGuarded => tElevatorUp, oReverseGuarded => tElevatorDown);
END_NETWORK
NETWORK 67 LD TITLE: "DONE NETWORK 44 (p3): Runtimeguard trayfiller"
  Mach1.GenFlags.StopDriveDirect S= RuntimeGuard_V5_1_100(Mach1_Alarms, (Mach1_AuxData.TrayfillerActive AND IDB_TrayFiller.oInfeedMotorFwd AND Mach1_AuxData.AllDrivesHomed), (Mach1_AuxData.TrayfillerActive AND IDB_TrayFiller.oInfeedMotorRev AND Mach1_AuxData.AllDrivesHomed), TRUE, T#4000MS, Mach1.GenFlags.StartFlag, Mach1_Alarms.Alm065, Mach1.GenFlags.MinorAlarm, Mach1_AuxData.IEC_TIMERS.RuntimeGuardInfeedConveyor, oForwardGuarded => LST_InputsOutputs.Q133_5_InfeedConv_Fwd, oReverseGuarded => LST_InputsOutputs.Q133_6_InfeedConv_Rev);
END_NETWORK
NETWORK 68 LD TITLE: "DONE NETWORK 44 (p4): Runtimeguard trayfiller"
  Mach1.GenFlags.StopDriveDirect S= RuntimeGuard_V5_1_100(Mach1_Alarms, (Mach1_AuxData.TrayfillerActive AND IDB_TrayFiller.oOutfeedMotorFwd AND Mach1_AuxData.AllDrivesHomed), NOT TRUE, TRUE, T#8500MS, Mach1.GenFlags.StartFlag, Mach1_Alarms.Alm066, Mach1.GenFlags.MinorAlarm, Mach1_AuxData.IEC_TIMERS.RuntimeGuardOutfeedConveyor, oForwardUnguarded => tBool, oForwardGuarded => LST_InputsOutputs.Q133_7_OutfeedConv_Fwd, oReverseUnguarded => tBool, oReverseGuarded => tBool);
END_NETWORK
NETWORK 69 LD TITLE: "DONE NETWORK 45: Elevator: profinet vs IO"
  LET g21 := (tElevatorUp OR tElevatorDown);
  Mach1_Data.Drives.ElevatorATF.Control.StartAuto := g21;
  LET en1 := g21;
  IF en1 THEN Mach1_Data.Drives.ElevatorATF.Control.AutoSpeed := MOVE(30); END_IF
  Mach1_Data.Drives.ElevatorATF.Control.Reverse := (g21 AND tElevatorDown);
END_NETWORK
NETWORK 70 LD TITLE: "DONE NETWORK 46 (p1): Alarms trayfiller"
  Mach1.GenFlags.StopDriveDirect S= Alarms_V5_1_100(Mach1_Alarms, (Mach1_AuxData.TrayfillerActive AND Mach1.GenFlags.DelayAfterEmergStop AND Mach1.GenFlags.DelayAfterSTO AND NOT LST_InputsOutputs.I132_0_Thermal_guards_OK AND (Mach1_AuxData.AllDrivesHomed OR NOT Mach1_AuxData.MIDS_Active)), Mach1.GenFlags.StartFlag, Mach1_Alarms.Alm005, Mach1.GenFlags.MinorAlarm);
END_NETWORK
NETWORK 71 LD TITLE: "DONE NETWORK 46 (p2): Alarms trayfiller"
  Mach1.GenFlags.StopDriveDirect S= Alarms_V5_1_100(Mach1_Alarms, (Mach1_AuxData.TrayfillerActive AND Trayfiller_Data.Alarms.AlmInpusherBlocked AND (Mach1_AuxData.AllDrivesHomed OR NOT Mach1_AuxData.MIDS_Active)), Mach1.GenFlags.StartFlag, Mach1_Alarms.Alm059, Mach1.GenFlags.MinorAlarm);
END_NETWORK
NETWORK 72 LD TITLE: "DONE NETWORK 46 (p3): Alarms trayfiller"
  Mach1.GenFlags.StopDriveDirect S= Alarms_V5_1_100(Mach1_Alarms, (Mach1_AuxData.TrayfillerActive AND (Trayfiller_Data.Alarms.AlmTrayPosition OR Trayfiller_Data.Alarms.AlmTrayInfeeding) AND Mach1_AuxData.AllDrivesHomed), TRUE, Mach1_Alarms.Alm060, Mach1.GenFlags.MinorAlarm);
END_NETWORK
NETWORK 73 LD TITLE: "DONE NETWORK 46 (p4): Alarms trayfiller"
  Mach1.GenFlags.StopDriveDirect S= Alarms_V5_1_100(Mach1_Alarms, (Mach1_AuxData.TrayfillerActive AND Trayfiller_Data.Alarms.AlmLightCurtainInpusher AND (Mach1_AuxData.AllDrivesHomed OR NOT Mach1_AuxData.MIDS_Active)), Mach1.GenFlags.StartFlag, Mach1_Alarms.Alm061, Mach1.GenFlags.MinorAlarm);
END_NETWORK
NETWORK 74 LD TITLE: "DONE NETWORK 46 (p5): Alarms trayfiller"
  Alarms_V5_1_100(Mach1_Alarms, (Mach1_AuxData.TrayfillerActive AND Trayfiller_Data.Alarms.WrnChangeTray AND (Mach1_AuxData.AllDrivesHomed OR NOT Mach1_AuxData.MIDS_Active)), TRUE, Mach1_Alarms.Alm075, Mach1.GenFlags.Warning);
END_NETWORK
NETWORK 75 LD TITLE: "DONE NETWORK 46 (p6): Alarms trayfiller"
  Alarms_V5_1_100(Mach1_Alarms, (Mach1_AuxData.TrayfillerActive AND Trayfiller_Data.Alarms.AlmOutfeedFull AND (Mach1_AuxData.AllDrivesHomed OR NOT Mach1_AuxData.MIDS_Active)), TRUE, Mach1_Alarms.Alm062, Mach1.GenFlags.MinorAlarm);
END_NETWORK
NETWORK 76 LD TITLE: "DONE NETWORK 46 (p7): Alarms trayfiller"
  Alarms_V5_1_100(Mach1_Alarms, (Mach1_AuxData.TrayfillerActive AND Trayfiller_Data.Alarms.AlmOutfeeding AND (Mach1_AuxData.AllDrivesHomed OR NOT Mach1_AuxData.MIDS_Active)), TRUE, Mach1_Alarms.Alm063, Mach1.GenFlags.MinorAlarm);
END_NETWORK
NETWORK 77 LD TITLE: "DONE NETWORK 46 (p8): Alarms trayfiller"
  Mach1.GenFlags.StopDriveDirect S= Alarms_V5_1_100(Mach1_Alarms, (Mach1_AuxData.TrayfillerActive AND Trayfiller_Data.Alarms.AlmLightCurtainElevator AND (Mach1_AuxData.AllDrivesHomed OR NOT Mach1_AuxData.MIDS_Active)), TRUE, Mach1_Alarms.Alm064, Mach1.GenFlags.MinorAlarm);
END_NETWORK
NETWORK 78 LD TITLE: "DONE NETWORK 46 (p9): Alarms trayfiller"
  Mach1.GenFlags.StopDriveDirect S= (Mach1_AuxData.AllDrivesHomed AND Mach1_AuxData.TrayfillerActive AND NOT Trayfiller_Data.commInterface.Permission);
END_NETWORK
NETWORK 79 LD TITLE: "TODO NETWORK 47 (p1):Greasing system"
END_NETWORK
NETWORK 80 LD TITLE: "DONE NETWORK 47 (p2): Greasing system"
  Mach1.GenFlags.StopDriveDirect S= Alarms_V5_1_100(Mach1_Alarms, (Mach1.GenFlags.DelayAfterEmergStop AND tLowLevel), TRUE, Mach1_Alarms.Alm078, Mach1.GenFlags.Warning);
END_NETWORK
NETWORK 81 LD TITLE: "DONE NETWORK 48: Alarm: Greasing system"
  Mach1.GenFlags.StopDriveDirect S= Alarms_V5_1_100(Mach1_Alarms, (Mach1.GenFlags.DelayAfterEmergStop AND tErrorRuntimeGreasingSystem), Mach1.GenFlags.StartFlag, Mach1_Alarms.Alm067, Mach1.GenFlags.MinorAlarm);
END_NETWORK
NETWORK 82 LD TITLE: "DONE NETWORK 49: State of the machine"
  LET g22 := TRUE;
  LET en1 := (g22 AND (Mach1.GenFlags.MajorAlarm OR Mach1.GenFlags.MinorAlarm));
  IF en1 THEN HMI_Var.Mach1.Status := MOVE(0); END_IF
  tAlarmSL := en1;
  LET g23 := (g22 AND NOT Mach1.GenFlags.MajorAlarm AND NOT Mach1.GenFlags.MinorAlarm);
  LET en2 := (g23 AND Mach1.GenFlags.Warning);
  IF en2 THEN HMI_Var.Mach1.Status := MOVE(1); END_IF
  tWarningSL := en2;
  LET g24 := (g23 AND NOT Mach1.GenFlags.Warning);
  LET en3 := (g24 AND NOT Mach1.GenFlags.RunMan AND NOT Mach1.GenFlags.RunAuto);
  IF en3 THEN HMI_Var.Mach1.Status := MOVE(2); END_IF
  tStandbySL := en3;
  LET en4 := (g24 AND (Mach1.GenFlags.RunMan OR Mach1.GenFlags.RunAuto));
  IF en4 THEN HMI_Var.Mach1.Status := MOVE(3); END_IF
  tRunningSL := en4;
END_NETWORK
NETWORK 83 LD TITLE: "TODO NETWORK 50: SL Alarmlamp"
  LET g25 := TRUE;
  LST_InputsOutputs.Q100_2_Pilot_light_Alarm_red_ := (g25 AND tAlarmlamp AND tAlarmSL);
  LST_InputsOutputs.Q100_1_Pilot_light_Alarm_orange_ := (g25 AND tAlarmlamp AND tWarningSL);
  LST_InputsOutputs.Q100_0_Pilot_light_Alarm_green_ := (g25 AND ((tAlarmlamp AND tStandbySL) OR tRunningSL));
END_NETWORK
NETWORK 84 LD TITLE: "TODO NETWORK 51: SL Alarmlamp Buzzer"
END_NETWORK

END_PROGRAM

(* ---- SMC_BitsToBytes.prg ---- *)
PROGRAM SMC_BitsToBytes
VAR
END_VAR

LST_InputsOutputs.SMC_B0.0:= BOOL_TO_BIT( PneumValveTerminalSMC.Pos1A);
LST_InputsOutputs.SMC_B0.1:= BOOL_TO_BIT( PneumValveTerminalSMC.Pos1B);
LST_InputsOutputs.SMC_B0.2:= BOOL_TO_BIT( PneumValveTerminalSMC.Pos2A);
LST_InputsOutputs.SMC_B0.3:= BOOL_TO_BIT( PneumValveTerminalSMC.Pos2B);
LST_InputsOutputs.SMC_B0.4:= BOOL_TO_BIT( PneumValveTerminalSMC.Pos3A);
LST_InputsOutputs.SMC_B0.5:= BOOL_TO_BIT( PneumValveTerminalSMC.Pos3B);
LST_InputsOutputs.SMC_B0.6:= BOOL_TO_BIT( PneumValveTerminalSMC.Pos4A);
LST_InputsOutputs.SMC_B0.7:= BOOL_TO_BIT( PneumValveTerminalSMC.Pos4B);

LST_InputsOutputs.SMC_B1.0:= BOOL_TO_BIT( PneumValveTerminalSMC.Pos5A);
LST_InputsOutputs.SMC_B1.1:= BOOL_TO_BIT( PneumValveTerminalSMC.Pos5B);
LST_InputsOutputs.SMC_B1.2:= BOOL_TO_BIT( PneumValveTerminalSMC.Pos6A);
LST_InputsOutputs.SMC_B1.3:= BOOL_TO_BIT( PneumValveTerminalSMC.Pos6B);
LST_InputsOutputs.SMC_B1.4:= BOOL_TO_BIT( PneumValveTerminalSMC.Pos7A);
LST_InputsOutputs.SMC_B1.5:= BOOL_TO_BIT( PneumValveTerminalSMC.Pos7B);
LST_InputsOutputs.SMC_B1.6:= BOOL_TO_BIT( PneumValveTerminalSMC.Pos8A);
LST_InputsOutputs.SMC_B1.7:= BOOL_TO_BIT( PneumValveTerminalSMC.Pos8B);

LST_InputsOutputs.SMC_B2.0:= BOOL_TO_BIT( PneumValveTerminalSMC.Pos9A);
LST_InputsOutputs.SMC_B2.1:= BOOL_TO_BIT( PneumValveTerminalSMC.Pos9B);
LST_InputsOutputs.SMC_B2.2:= BOOL_TO_BIT( PneumValveTerminalSMC.Pos10A);
LST_InputsOutputs.SMC_B2.3:= BOOL_TO_BIT( PneumValveTerminalSMC.Pos10B);
LST_InputsOutputs.SMC_B2.4:= BOOL_TO_BIT( PneumValveTerminalSMC.Pos11A);
LST_InputsOutputs.SMC_B2.5:= BOOL_TO_BIT( PneumValveTerminalSMC.Pos11B);
LST_InputsOutputs.SMC_B2.6:= BOOL_TO_BIT( PneumValveTerminalSMC.Pos12A);
LST_InputsOutputs.SMC_B2.7:= BOOL_TO_BIT( PneumValveTerminalSMC.Pos12B);
(*
LST_InputsOutputs.SMC_B3.0:= BOOL_TO_BIT( PneumValveTerminalSMC.Pos13A);
LST_InputsOutputs.SMC_B3.1:= BOOL_TO_BIT( PneumValveTerminalSMC.Pos13B);
LST_InputsOutputs.SMC_B3.2:= BOOL_TO_BIT( PneumValveTerminalSMC.Pos14A);
LST_InputsOutputs.SMC_B3.3:= BOOL_TO_BIT( PneumValveTerminalSMC.Pos14B);
LST_InputsOutputs.SMC_B3.4:= BOOL_TO_BIT( PneumValveTerminalSMC.Pos15A);
LST_InputsOutputs.SMC_B3.5:= BOOL_TO_BIT( PneumValveTerminalSMC.Pos15B);
LST_InputsOutputs.SMC_B3.6:= BOOL_TO_BIT( PneumValveTerminalSMC.Pos16A);
LST_InputsOutputs.SMC_B3.7:= BOOL_TO_BIT( PneumValveTerminalSMC.Pos16B);
*)

END_PROGRAM

(* ---- SMC_BytesToBits.prg ---- *)
PROGRAM SMC_BytesToBits
VAR
END_VAR

LST_InputsOutputs.SMC_B0.0:= BOOL_TO_BIT( PneumValveTerminalSMC.Pos1A);
LST_InputsOutputs.SMC_B0.1:= BOOL_TO_BIT( PneumValveTerminalSMC.Pos1B);
LST_InputsOutputs.SMC_B0.2:= BOOL_TO_BIT( PneumValveTerminalSMC.Pos2A);
LST_InputsOutputs.SMC_B0.3:= BOOL_TO_BIT( PneumValveTerminalSMC.Pos2B);
LST_InputsOutputs.SMC_B0.4:= BOOL_TO_BIT( PneumValveTerminalSMC.Pos3A);
LST_InputsOutputs.SMC_B0.5:= BOOL_TO_BIT( PneumValveTerminalSMC.Pos3B);
LST_InputsOutputs.SMC_B0.6:= BOOL_TO_BIT( PneumValveTerminalSMC.Pos4A);
LST_InputsOutputs.SMC_B0.7:= BOOL_TO_BIT( PneumValveTerminalSMC.Pos4B);

LST_InputsOutputs.SMC_B1.0:= BOOL_TO_BIT( PneumValveTerminalSMC.Pos5A);
LST_InputsOutputs.SMC_B1.1:= BOOL_TO_BIT( PneumValveTerminalSMC.Pos5A);
LST_InputsOutputs.SMC_B1.2:= BOOL_TO_BIT( PneumValveTerminalSMC.Pos6A);
LST_InputsOutputs.SMC_B1.3:= BOOL_TO_BIT( PneumValveTerminalSMC.Pos6B);
LST_InputsOutputs.SMC_B1.4:= BOOL_TO_BIT( PneumValveTerminalSMC.Pos7A);
LST_InputsOutputs.SMC_B1.5:= BOOL_TO_BIT( PneumValveTerminalSMC.Pos7B);
LST_InputsOutputs.SMC_B1.6:= BOOL_TO_BIT( PneumValveTerminalSMC.Pos8A);
LST_InputsOutputs.SMC_B1.7:= BOOL_TO_BIT( PneumValveTerminalSMC.Pos8B);

LST_InputsOutputs.SMC_B2.0:= BOOL_TO_BIT( PneumValveTerminalSMC.Pos9A);
LST_InputsOutputs.SMC_B2.1:= BOOL_TO_BIT( PneumValveTerminalSMC.Pos9B);
LST_InputsOutputs.SMC_B2.2:= BOOL_TO_BIT( PneumValveTerminalSMC.Pos10A);
LST_InputsOutputs.SMC_B2.3:= BOOL_TO_BIT( PneumValveTerminalSMC.Pos10B);
LST_InputsOutputs.SMC_B2.4:= BOOL_TO_BIT( PneumValveTerminalSMC.Pos11A);
LST_InputsOutputs.SMC_B2.5:= BOOL_TO_BIT( PneumValveTerminalSMC.Pos11B);
LST_InputsOutputs.SMC_B2.6:= BOOL_TO_BIT( PneumValveTerminalSMC.Pos12A);
LST_InputsOutputs.SMC_B2.7:= BOOL_TO_BIT( PneumValveTerminalSMC.Pos12B);
(*
SMC_B3.0:= BOOL_TO_BIT( PneumValveTerminalSMC.Pos13A);
SMC_B3.1:= BOOL_TO_BIT( PneumValveTerminalSMC.Pos13B);
SMC_B3.2:= BOOL_TO_BIT( PneumValveTerminalSMC.Pos14A);
SMC_B3.3:= BOOL_TO_BIT( PneumValveTerminalSMC.Pos14B);
SMC_B3.4:= BOOL_TO_BIT( PneumValveTerminalSMC.Pos15A);
SMC_B3.5:= BOOL_TO_BIT( PneumValveTerminalSMC.Pos15B);
SMC_B3.6:= BOOL_TO_BIT( PneumValveTerminalSMC.Pos16A);
SMC_B3.7:= BOOL_TO_BIT( PneumValveTerminalSMC.Pos16B);
*)

END_PROGRAM

(* ---- Status_ForceOutputs.prg ---- *)
PROGRAM Status_ForceOutputs
VAR
END_VAR

NETWORK 0 LD
  LET g9 := TRUE;
  LET en1 := g9;
  IF en1 THEN LST_InputsOutputs.Serv_IB100 := MOVE(%IB26); END_IF
  LET en2 := g9;
  IF en2 THEN LST_InputsOutputs.Serv_IB101 := MOVE(%IB27); END_IF
END_NETWORK
NETWORK 1 LD
  LET g13 := TRUE;
  LET en1 := g13;
  IF en1 THEN LST_InputsOutputs.Serv_IB132 := MOVE(%IB370); END_IF
  LET en2 := g13;
  IF en2 THEN LST_InputsOutputs.Serv_IB133 := MOVE(%IB371); END_IF
  LET en3 := g13;
  IF en3 THEN LST_InputsOutputs.Serv_IB136 := MOVE(%IB372); END_IF
  LET en4 := g13;
  IF en4 THEN LST_InputsOutputs.Serv_IB137 := MOVE(%IB373); END_IF
END_NETWORK
NETWORK 2 LD
  LET en1 := HMI_Var.ForceOutputs;
  IF en1 THEN ForceOutput(); END_IF
END_NETWORK
NETWORK 3 LD
  LET en1 := NOT HMI_Var.ForceOutputs;
  IF en1 THEN ForceOutput_1(); END_IF
END_NETWORK
NETWORK 4 LD
END_NETWORK

END_PROGRAM
